(* IEC 61131-3 sources: daoli-st-library/DL_MathData (part 3) *)

(* ---- FC_DL_InterpSegmentWeight.st ---- *)
(*==============================================================================
 * 组件名称 (Component)  : FC_DL_InterpSegmentWeight
 * 所属子库 (Sublibrary) : DL_MathData
 * 当前版本 (Version)    : 1.0.0
 * 兼容性   (Platform)   : CODESYS 3.5+ / TwinCAT 3 / 汇川 InoProShop / 施耐德 Machine Expert
 *                         仅依赖 IEC 61131-3 标准数学（ABS / MIN / MAX），零厂商私有库
 * 功能描述 (Function)   : 段内权重计算：给定升序节点表与查询点，返回相邻两点的
 *                         **加权系数对** (fWLeft, fWRight)，满足 fWLeft + fWRight = 1：
 *                           fWRight = (fXin - afX[i]) / (afX[i+1] - afX[i])
 *                           fWLeft  = 1 - fWRight
 *                         调用方据此自行取 Y（若只有 Y 单表，可算 y = wl*y_i + wr*y_{i+1}），
 *                         也可用于多表共享同一权重（同一 X 上插值多条曲线，
 *                         避免重复定位，性能与一致性双收益）。
 *                         v = wl*v_i + wr*v_{i+1} 与线性插值严格等价（权重和为 1 保证无偏）。
 * 接口     (Interface)  : 输入 afX 升序节点表 [X 单位]、iCount 有效点数 [个]（2..32）、
 *                         fXin 查询点 [X 单位]；
 *                         输出 iSeg 区间左端下标、fWLeft 左节点权重 [0..1]、
 *                         fWRight 右节点权重 [0..1]、bClamped 越界钳位回执、
 *                         eErrCode（E_DL_InterpWgtErr）；
 *                         返回值 = bValid 权重可信标志（TRUE = 两权重可信）。
 * 边界     (Boundary)   : ① 属主边界：只给权重，**不取 Y 值**（取值由调用方组合，
 *                         这是本件与 InterpHoldLast / TwoPointSlope 的本质分工）。
 *                         ② 点数域闸 2..32；越域 → 故障级 eBadCount。
 *                         ③ 非有限双判：查询点 + 全部表元素逐项枚举。
 *                         ④ 段宽近似零 → fWLeft=1.0、fWRight=0.0 并置信息级 eDegenerateSeg
 *                         （权重仍满足和为 1，调用方无需特判；除零被完全规避）。
 *                         ⑤ 越界钳位：fXin 超出 [afX[1], afX[iCount]] → 钳到端段端点，
 *                         权重退化为 (1,0) 或 (0,1)，bClamped=TRUE，不外推。
 *                         ⑥ 权重和复检：|fWLeft + fWRight - 1| < 1E-9，违反 → 故障级 eInternal
 *                         （结构性断言，防未来改动破坏无偏性）。
 *                         ⑦ 零全局耦合（无 GVL / VAR_EXTERNAL / 物理地址）。
 * 分工声明 (Scope)      : 与 `FC_DL_InterpHoldLast` 分工：那件直接给 Y（保持型），
 *                         本件只给权重（多表共享）；与 `FC_DL_TableIndexBinarySearch` 分工：
 *                         大表定位优先用那件，本件为线性扫描 + 权重输出件。
 * 来源标签 (Source Tag) : 原创实现（无外部代码引入）
 * 码表     (Codes)      : 本件不占用全局数字码位；出口为 BOOL + INT + 2×LREAL + BOOL +
 *                         本文件内定义 enum E_DL_InterpWgtErr（全库唯一）。
 * 红线自检 (Redline)    : R1 ✓ 零 GVL/VAR_EXTERNAL ｜ R2 ✓ 零 %I/%Q/%M ｜ R3 ✓ 纯 IEC 61131-3
 *                         R4 ✓ 点数域闸 + 全表非有限双判 + 段宽判零 + 权重和复检 ｜ R5 ✓ 声明逐行同行双语注释
 *                         R6 N/A（纯函数无状态机） ｜ R7 N/A（无实例调用）
 * 修订历史 (Revision)   : 2026-11-23  v1.0.0  R77 首版（批次 B3 · 序号 8）
 * 验收向量 (Acceptance) : ① afX=[0,10,20], iCount=3, fXin=5 → iSeg=1, fWRight=0.5,
 *                         fWLeft=0.5, bClamped=FALSE, eOk, TRUE；
 *                         ② afX 同上, fXin=15 → iSeg=2, fWRight=0.5, fWLeft=0.5；
 *                         ③ afX 同上, fXin=-3 → iSeg=1, fWLeft=1.0, fWRight=0.0, bClamped=TRUE；
 *                         ④ afX 同上, fXin=99 → iSeg=2, fWLeft=0.0, fWRight=1.0, bClamped=TRUE；
 *                         ⑤ afX=[0,0,20], fXin=0 → 退化段：fWLeft=1.0, fWRight=0.0, eDegenerateSeg。
 *==============================================================================*)

(*-----------------------------------------------------------------------------
 * 枚举: E_DL_InterpWgtErr（段内权重错误码，归属 DL_MathData，与本件同文件，全库唯一属主）
 *----------------------------------------------------------------------------*)
TYPE E_DL_InterpWgtErr :
(
    eOk            := 0,   // 信息级：权重计算完成 / Info: weights computed
    eDegenerateSeg := 1,   // 信息级：段宽近似零，权重退化为 1/0 / Info: degenerate segment, weights 1 and 0
    eBadCount      := 2,   // 故障级：点数越域 / Fault: point count out of domain
    eNonFinite     := 3,   // 故障级：查询点或表元素非有限 / Fault: query or table entry non-finite
    eTableNotAsc   := 4,   // 故障级：表不满足升序约定 / Fault: table violates ascending contract
    eInternal      := 9    // 故障级：权重和偏离 1，无偏性被破坏 / Fault: weight sum deviates from one
);
END_TYPE

FUNCTION FC_DL_InterpSegmentWeight : BOOL
VAR_INPUT
    afX    : ARRAY[1..32] OF LREAL;  // 升序节点表 [X 单位] / Ascending node table in X
    iCount : INT;                    // 有效点数（2..32） [个] / Valid point count, 2..32
    fXin   : LREAL;                  // 查询点 [X 单位] / Query value in X
END_VAR
VAR_OUTPUT
    iSeg     : INT;    // 区间左端下标（1..iCount-1） [-] / Segment left index
    fWLeft   : LREAL;  // 左节点权重 [0..1] [-] / Left node weight
    fWRight  : LREAL;  // 右节点权重 [0..1] [-] / Right node weight
    bClamped : BOOL;   // 越界钳位回执 [-] / Out-of-range clamp receipt
    eErrCode : E_DL_InterpWgtErr; // 错误码出口 [-] / Error code outlet
END_VAR
VAR
    _i       : INT;    // 循环下标 [-] / Loop index
    _iSeg    : INT;    // 命中区间下标 [-] / Hit segment index
    _bFound  : BOOL;   // 区间命中标志 [-] / Segment found flag
    _bNonFin : BOOL;   // 非有限标志 [-] / Non-finite flag
    _fDen    : LREAL;  // 段宽（分母） [X 单位] / Segment width denominator
    _fWr     : LREAL;  // 右权重（未钳位） [-] / Raw right weight
    _fSum    : LREAL;  // 权重和（复检用） [-] / Weight sum for recheck
END_VAR
VAR CONSTANT
    DL_IWC_CNT_MIN : INT := 2;        // 点数下限 [个] / Count lower bound
    DL_IWC_CNT_MAX : INT := 32;       // 点数上限（数组容量） [个] / Count upper bound
    DL_IWC_TINY    : LREAL := 1.0E-9; // 段宽近似零阈值 [X 单位] / Degenerate segment threshold
    DL_IWC_ZERO    : LREAL := 0.0;    // 零与权重下限 [-] / Zero and weight lower bound
    DL_IWC_ONE     : LREAL := 1.0;    // 权重上限与无偏基准 [-] / Weight upper bound and unbiasedness base
END_VAR

(* —— 段 0：出口预置安全值（权重预置为「全取左端」，恒满足和为 1） —— *)
FC_DL_InterpSegmentWeight := FALSE;                // 返回值预置无效 / Return preset invalid
iSeg     := 0;                                     // 下标哨兵 / Index sentinel
fWLeft   := DL_IWC_ONE;                            // 左权重哨兵 1（最保守：全取左端） / Left weight sentinel
fWRight  := DL_IWC_ZERO;                           // 右权重哨兵 0 / Right weight sentinel
bClamped := FALSE;                                 // 钳位回执预置否 / Clamp receipt preset false
eErrCode := E_DL_InterpWgtErr.eBadCount;           // 预置最严码 / Preset strictest code

(* —— 段 1：点数域闸 —— *)
IF (iCount < DL_IWC_CNT_MIN) OR (iCount > DL_IWC_CNT_MAX) THEN
    RETURN;
END_IF

(* —— 段 2：非有限域闸（查询点 + 全部表元素逐项枚举） —— *)
_bNonFin := (fXin <> fXin) OR ((fXin - fXin) <> DL_IWC_ZERO);
_i := 1;
WHILE _i <= iCount DO
    IF (afX[_i] <> afX[_i]) OR ((afX[_i] - afX[_i]) <> DL_IWC_ZERO) THEN
        _bNonFin := TRUE;
    END_IF
    _i := _i + 1;
END_WHILE
IF _bNonFin THEN
    eErrCode := E_DL_InterpWgtErr.eNonFinite;
    RETURN;
END_IF

(* —— 段 3：下越界钳位（权重退化 1/0） —— *)
IF fXin <= afX[1] THEN
    iSeg     := 1;
    fWLeft   := DL_IWC_ONE;
    fWRight  := DL_IWC_ZERO;
    bClamped := TRUE;
    eErrCode := E_DL_InterpWgtErr.eOk;
    FC_DL_InterpSegmentWeight := TRUE;
    RETURN;
END_IF

(* —— 段 4：上越界钳位（权重退化 0/1） —— *)
IF fXin >= afX[iCount] THEN
    iSeg     := iCount - 1;
    fWLeft   := DL_IWC_ZERO;
    fWRight  := DL_IWC_ONE;
    bClamped := TRUE;
    eErrCode := E_DL_InterpWgtErr.eOk;
    FC_DL_InterpSegmentWeight := TRUE;
    RETURN;
END_IF

(* —— 段 5：区间定位（升序：afX[i] <= fXin <= afX[i+1]） —— *)
_i      := 1;
_bFound := FALSE;
_iSeg   := 1;
WHILE (_i < iCount) AND (NOT _bFound) DO
    IF (fXin >= afX[_i]) AND (fXin <= afX[_i + 1]) THEN
        _bFound := TRUE;
        _iSeg   := _i;
    ELSE
        _i := _i + 1;
    END_IF
END_WHILE
IF NOT _bFound THEN
    eErrCode := E_DL_InterpWgtErr.eTableNotAsc;    // 未命中：表不升序 / Not found: table not ascending
    RETURN;
END_IF

(* —— 段 6：升序复检 + 段宽判零后计算权重 —— *)
IF afX[_iSeg + 1] < afX[_iSeg] THEN
    eErrCode := E_DL_InterpWgtErr.eTableNotAsc;    // 端点倒序 / Endpoints reversed
    RETURN;
END_IF
_fDen := afX[_iSeg + 1] - afX[_iSeg];              // 段宽 / Segment width
IF ABS(_fDen) < DL_IWC_TINY THEN
    fWLeft   := DL_IWC_ONE;                        // 退化段：全取左端 / Degenerate: all to left
    fWRight  := DL_IWC_ZERO;
    eErrCode := E_DL_InterpWgtErr.eDegenerateSeg;  // 信息级码 / Info code
ELSE
    _fWr     := (fXin - afX[_iSeg]) / _fDen;       // 右权重 / Right weight
    fWRight  := MIN(MAX(_fWr, DL_IWC_ZERO), DL_IWC_ONE);      // 显式约束 0..1 / Constrain 0..1
    fWLeft   := DL_IWC_ONE - fWRight;              // 左权重 = 1 - 右权重（无偏性构造） / Left weight
    eErrCode := E_DL_InterpWgtErr.eOk;             // 信息级成功 / Info success
END_IF
iSeg := _iSeg;

(* —— 段 7：权重和无偏性复检（结构性断言） —— *)
_fSum := fWLeft + fWRight;                         // 权重和 / Weight sum
IF ABS(_fSum - DL_IWC_ONE) > DL_IWC_TINY THEN
    fWLeft   := DL_IWC_ONE;                        // 复检失败：回最保守权重 / Recheck failed: conservative weights
    fWRight  := DL_IWC_ZERO;
    iSeg     := 0;
    eErrCode := E_DL_InterpWgtErr.eInternal;       // 故障级：内部不一致 / Fault: internal inconsistency
    RETURN;
END_IF

FC_DL_InterpSegmentWeight := TRUE;                 // 权重可信 / Weights trustworthy

END_FUNCTION

(* ---- FC_DL_InterpTwoPointSlope.st ---- *)
(*==============================================================================
 * 组件名称 (Component)  : FC_DL_InterpTwoPointSlope
 * 所属子库 (Sublibrary) : DL_MathData
 * 当前版本 (Version)    : 1.0.0
 * 兼容性   (Platform)   : CODESYS 3.5+ / TwinCAT 3 / 汇川 InoProShop / 施耐德 Machine Expert
 *                         仅依赖 IEC 61131-3 标准数学（ABS），零厂商私有库
 * 功能描述 (Function)   : 两点定斜率线性插值 / 受限外推。
 *                           k  = (y2 - y1) / (x2 - x1)                 —— 由两点确定
 *                           y  = y1 + k × (xin - x1)                    —— 通用式（插值外推同一式）
 *                         外推保护：外推距离 = |xin - 近端节点 X|，若超过 fMaxExtrap
 *                         （默认 0.0 = 禁止外推，仅区间内插值），则把 xin 钳到
 *                         「近端节点 ± fMaxExtrap」后再取值，并置 bExtrapolated
 *                         与信息级 eExtrapClamped。**钳位的是 xin 而非 y**，
 *                         这样斜率信息仍可复用（调用方可用 fSlope 自行延续）。
 * 接口     (Interface)  : 输入 fX1/fY1 节点 1、fX2/fY2 节点 2、fXin 查询点、
 *                         fMaxExtrap 允许的最大外推距离 [X 单位，0 = 禁止外推]；
 *                         输出 fYout 结果 [Y 单位]、fSlope 斜率 [Y/X]、
 *                         bExtrapolated 是否发生外推、eErrCode（E_DL_InterpSlopeErr）；
 *                         返回值 = bValid 结果可信标志（TRUE = fYout 可信）。
 * 边界     (Boundary)   : ① 属主边界：只做两点定斜率，不做多点表遍历、不做曲线拟合。
 *                         ② 全浮点入参（7 个）非有限双判，逐一枚举。
 *                         ③ 两点 X 重合（|x2-x1| < 1E-9）→ 故障级 eDegenerateNodes
 *                         （斜率无定义，禁止除零；**先判零后除**）。
 *                         ④ fMaxExtrap < 0 → 故障级 eBadParam（负外推距离无意义）。
 *                         ⑤ fMaxExtrap = 0 表示禁止外推：xin 越界即钳到节点 X，结果 = 端点 Y。
 *                         ⑥ 零全局耦合（无 GVL / VAR_EXTERNAL / 物理地址）。
 * 分工声明 (Scope)      : 与 `FC_DL_InterpLogLinear` 分工：对数域归那件、线性域归本件；
 *                         与 `FC_DL_InterpHoldLast` 分工：保持型（不外推只保持）归那件。
 * 来源标签 (Source Tag) : 原创实现（无外部代码引入）
 * 码表     (Codes)      : 本件不占用全局数字码位；出口为 BOOL + 2×LREAL + BOOL +
 *                         本文件内定义 enum E_DL_InterpSlopeErr（全库唯一）。
 * 红线自检 (Redline)    : R1 ✓ 零 GVL/VAR_EXTERNAL ｜ R2 ✓ 零 %I/%Q/%M ｜ R3 ✓ 纯 IEC 61131-3
 *                         R4 ✓ 全入参非有限双判 + 两点 X 重合判零（除零防护）+ 外推距离上限 ｜ R5 ✓ 声明逐行同行双语注释
 *                         R6 N/A（纯函数无状态机） ｜ R7 N/A（无实例调用）
 * 修订历史 (Revision)   : 2026-11-23  v1.0.0  R77 首版（批次 B3 · 序号 4）
 * 验收向量 (Acceptance) : ① fX1=0, fY1=0, fX2=10, fY2=100, fXin=5, fMaxExtrap=0 → k=10,
 *                         fYout=50.0, bExtrapolated=FALSE, eOk；
 *                         ② 同上, fXin=12, fMaxExtrap=5 → 外推 2 <= 5 → fYout=120.0, eExtrapolated；
 *                         ③ 同上, fXin=20, fMaxExtrap=5 → 钳 xin 到 15 → fYout=150.0, eExtrapClamped；
 *                         ④ fX1=fX2=5 → 返回 FALSE, fYout=0, eDegenerateNodes；
 *                         ⑤ fXin=0, fMaxExtrap=0 → fYout=0.0（左端外推钳到 x1）。
 *==============================================================================*)

(*-----------------------------------------------------------------------------
 * 枚举: E_DL_InterpSlopeErr（两点定斜率插值错误码，归属 DL_MathData，与本件同文件，全库唯一属主）
 *----------------------------------------------------------------------------*)
TYPE E_DL_InterpSlopeErr :
(
    eOk             := 0,   // 信息级：区间内插值 / Info: in-range interpolation
    eExtrapolated   := 1,   // 信息级：受限外推（未超限） / Info: bounded extrapolation within limit
    eExtrapClamped  := 2,   // 信息级：外推超限已钳位 / Info: extrapolation clamped to limit
    eDegenerateNodes:= 3,   // 故障级：两点 X 重合，斜率无定义 / Fault: coincident X, undefined slope
    eBadParam       := 4,   // 故障级：外推距离参数为负 / Fault: negative extrapolation distance
    eNonFinite      := 5    // 故障级：入参非有限 / Fault: non-finite input
);
END_TYPE

FUNCTION FC_DL_InterpTwoPointSlope : BOOL
VAR_INPUT
    fX1        : LREAL;  // 节点 1 的 X [X 单位] / Node one X
    fY1        : LREAL;  // 节点 1 的 Y [Y 单位] / Node one Y
    fX2        : LREAL;  // 节点 2 的 X [X 单位] / Node two X
    fY2        : LREAL;  // 节点 2 的 Y [Y 单位] / Node two Y
    fXin       : LREAL;  // 查询点 X [X 单位] / Query X
    fMaxExtrap : LREAL;  // 允许的最大外推距离（0 = 禁止外推） [X 单位] / Max extrapolation distance, zero forbids
END_VAR
VAR_OUTPUT
    fYout         : LREAL;  // 插值 / 外推结果 [Y 单位] / Interpolated or extrapolated result
    fSlope        : LREAL;  // 两点定出的斜率 [Y/X 单位比] / Slope determined by the two nodes
    bExtrapolated : BOOL;   // 是否发生外推 [-] / Whether extrapolation occurred
    eErrCode      : E_DL_InterpSlopeErr; // 错误码出口 [-] / Error code outlet
END_VAR
VAR
    _bNonFin : BOOL;   // 入参非有限标志 [-] / Non-finite input flag
    _fDx     : LREAL;  // X 方向增量 [X 单位] / X increment
    _fOut    : LREAL;  // 外推距离（带符号） [X 单位] / Signed extrapolation distance
    _fXUse   : LREAL;  // 钳位后实际使用的 X [-] / Actually used X after clamping
    _fLo     : LREAL;  // 允许区间左界 [X 单位] / Allowed lower bound
    _fHi     : LREAL;  // 允许区间右界 [X 单位] / Allowed upper bound
END_VAR
VAR CONSTANT
    DL_ITS_ZERO : LREAL := 0.0;     // 零基准 [-] / Zero base
    DL_ITS_TINY : LREAL := 1.0E-9;  // 两点 X 重合阈值 [X 单位] / Coincident X threshold
END_VAR

(* —— 段 0：出口预置安全值 —— *)
FC_DL_InterpTwoPointSlope := FALSE;                // 返回值预置无效 / Return preset invalid
fYout         := DL_ITS_ZERO;                      // 结果哨兵 0 / Result sentinel
fSlope        := DL_ITS_ZERO;                      // 斜率哨兵 0 / Slope sentinel
bExtrapolated := FALSE;                            // 外推标志预置否 / Extrapolation preset false
eErrCode      := E_DL_InterpSlopeErr.eBadParam;    // 预置最严码 / Preset strictest code

(* —— 段 1：非有限域闸（6 个浮点入参逐一枚举） —— *)
_bNonFin := (fX1 <> fX1) OR ((fX1 - fX1) <> DL_ITS_ZERO);            // X1 非有限 / X1 non-finite
_bNonFin := _bNonFin OR (fY1 <> fY1) OR ((fY1 - fY1) <> DL_ITS_ZERO); // Y1 非有限 / Y1 non-finite
_bNonFin := _bNonFin OR (fX2 <> fX2) OR ((fX2 - fX2) <> DL_ITS_ZERO); // X2 非有限 / X2 non-finite
_bNonFin := _bNonFin OR (fY2 <> fY2) OR ((fY2 - fY2) <> DL_ITS_ZERO); // Y2 非有限 / Y2 non-finite
_bNonFin := _bNonFin OR (fXin <> fXin) OR ((fXin - fXin) <> DL_ITS_ZERO);       // 查询点非有限 / Query non-finite
_bNonFin := _bNonFin OR (fMaxExtrap <> fMaxExtrap) OR ((fMaxExtrap - fMaxExtrap) <> DL_ITS_ZERO); // 外推上限非有限
IF _bNonFin THEN
    eErrCode := E_DL_InterpSlopeErr.eNonFinite;    // 故障级码 / Fault-level code
    RETURN;
END_IF

(* —— 段 2：外推距离参数域闸（不得为负） —— *)
IF fMaxExtrap < DL_ITS_ZERO THEN
    eErrCode := E_DL_InterpSlopeErr.eBadParam;     // 故障级：参数非法 / Fault: illegal parameter
    RETURN;
END_IF

(* —— 段 3：两点 X 重合判零（先判零后做除法，R4 除零防护） —— *)
_fDx := fX2 - fX1;                                 // X 方向增量（分母） / X increment denominator
IF ABS(_fDx) < DL_ITS_TINY THEN
    eErrCode := E_DL_InterpSlopeErr.eDegenerateNodes;  // 故障级：斜率无定义 / Fault: undefined slope
    RETURN;                                        // 早退，杜绝除零 / Early exit, avoids division by zero
END_IF

(* —— 段 4：斜率计算 —— *)
fSlope := (fY2 - fY1) / _fDx;                      // k = dy / dx / Slope

(* —— 段 5：外推距离判定与钳位（钳 xin，不钳 y） —— *)
IF fXin < fX1 THEN
    _fOut := fX1 - fXin;                           // 左向外推距离（正数） / Left extrapolation distance
    IF _fOut > fMaxExtrap THEN
        _fXUse   := fX1 - fMaxExtrap;              // 钳到允许的最远点 / Clamp to farthest allowed point
        eErrCode := E_DL_InterpSlopeErr.eExtrapClamped;   // 信息级：超限钳位 / Info: clamped
    ELSE
        _fXUse   := fXin;                          // 未超限：原值使用 / Within limit: use as-is
        eErrCode := E_DL_InterpSlopeErr.eExtrapolated;    // 信息级：受限外推 / Info: bounded extrapolation
    END_IF
    bExtrapolated := TRUE;                         // 左向外推 / Left extrapolation
ELSIF fXin > fX2 THEN
    _fOut := fXin - fX2;                           // 右向外推距离（正数） / Right extrapolation distance
    IF _fOut > fMaxExtrap THEN
        _fXUse   := fX2 + fMaxExtrap;              // 钳到允许的最远点 / Clamp to farthest allowed point
        eErrCode := E_DL_InterpSlopeErr.eExtrapClamped;   // 信息级：超限钳位 / Info: clamped
    ELSE
        _fXUse   := fXin;                          // 未超限：原值使用 / Within limit: use as-is
        eErrCode := E_DL_InterpSlopeErr.eExtrapolated;    // 信息级：受限外推 / Info: bounded extrapolation
    END_IF
    bExtrapolated := TRUE;                         // 右向外推 / Right extrapolation
ELSE
    _fXUse        := fXin;                         // 区间内插值，无外推 / In-range interpolation
    bExtrapolated := FALSE;
    eErrCode      := E_DL_InterpSlopeErr.eOk;      // 信息级成功 / Info success
END_IF

(* —— 段 6：取值（插值与外推同一式） —— *)
fYout := fY1 + fSlope * (_fXUse - fX1);            // y = y1 + k*(x - x1)

(* —— 段 7：结果非有限复检兜底 —— *)
IF (fYout <> fYout) OR ((fYout - fYout) <> DL_ITS_ZERO) THEN
    fYout         := DL_ITS_ZERO;                  // 复检异常回哨兵 / Recheck failed: sentinel
    fSlope        := DL_ITS_ZERO;
    bExtrapolated := FALSE;
    eErrCode      := E_DL_InterpSlopeErr.eNonFinite;   // 故障级码 / Fault-level code
    RETURN;
END_IF

FC_DL_InterpTwoPointSlope := TRUE;                 // 结果有效 / Result valid

END_FUNCTION

(* ---- FC_DL_IntervalGapCalc.st ---- *)
(*
  ==================================================================
  组件名 Component  : FC_DL_IntervalGapCalc
  分类   Category   : DL_MathData
  前缀   Naming     : FC_DL_ ｜ b/n/u/f/t/e/st 类型前缀制（R265）
  码位   Code ID    : 16#0001_0665（故障级）
  版本   Version    : 1.0.0
  复杂度 Complexity  : 中
  功能   Purpose    : 两区间相离间隙计算：相离返回正间隙宽 [工程单位]，相接 /
                      重叠 / 包含返回 0 并带关系码；供工艺窗对撞分析、换型
                      死区校验、安全包络间距核算等调用方使用。
  开源溯源 Origin    : 西门子 LGF V5.3.0 Comparator 组「区间关系」分类事实
                      借鉴（只借骨不抄肉，与 R11 RangeOverlapCheck 同组既有
                      件互引）；间隙计算 clean-room，零代码复制。
  许可证 License    : MIT
  参考   Reference  : IEC 61131-3:2013 §6.6.1 比较 / MAX 语义
  平台   Platform   : 纯 IEC 61131-3（MAX / ABS / 比较），三平台通用
  依赖   Depends    : 无（零委托、零库件）
  分工声明 Split     : FC_DL_RangeOverlapCheck（五分支关系判定，输出重叠长度）
                      为姊妹件（互引）；本件为「间隙方向」补口：输出相离
                      间隙宽（RangeOverlapCheck 只输出重叠长度，相离时恒 0，
                      间隙量不可观测），两件口径差异显式声明（R216）。
  归属 Ownership     : E_DL_IntervalGap 属主为本文件（全库唯一定义，R264）；
                      引用件只引用不重声明。
  ------------------------------------------------------------------
  边界 Boundary     :
                      一 非有限闸（四个端点 + fEps 逐个点名，R272）：任一
                         非有限 → 故障级 0665 + 返回 eInvalid + fGap = 0 +
                         bValid = FALSE + 早退；
                      二 端点归一：每区间无序端点自动对调，保证下限 ≤ 上限；
                      三 fEps 域闸：负容差非法 → 按默认容差 1.0E-6 接管并
                         并入 0665 处置（与端点非有限出口同形：eInvalid +
                         fGap = 0 + bValid = FALSE，反证句见码表）；
                      四 判定次序写死：相离（正间隙 > fEps）→ 相接（端点
                         重合在容差内）→ 包含 → 部分重叠；相离必须先于
                         相接，相接必须先于重叠（次序不可调换，防多解）；
                      五 完全相等归入 eContained（含端点重合的包含）：相等
                         是包含的退化特例，间隙同为 0，出口无法区分（R90
                         不另立关系码，与 RangeOverlapCheck 的 eEqual 五分
                         支口径差异显式声明）；
                      六 fGap 返回前置非负钳位：舍入产生的微小负值钳到 0；
                      七 纯函数：无记忆量、无定时器、无边沿实例，每调用重算；
                      八 无除法、无循环、无数组访问；无全局、无外部变量、
                         无物理地址。
  错误码 Codes      :
    16#0001_0665【故障级】输入非有限（四端点 / fEps 为 NaN / ±Inf）或 fEps
                         为负（组态非法）
  码位反证 Note     :
    0665 合并「端点 / 容差非有限」与「fEps 为负」的理由：两场景出口组合完全
    相同（eInvalid、fGap = 0、bValid = FALSE、bError = TRUE），三组以内输出
    无法唯一还原该场景，按 R90 不另立码；eInvalid 关系码与 0665 分立：前者
    是返回值语义（关系不可判），后者是诊断码，通道不同不互斥。
  验收 Acceptance   :
    算法已证（脚本）：未跑 ｜ 编译器已证（三平台）：未跑
    V1 相离：A = [0, 10]、B = [20, 30] → eDisjoint、fGap = 10.0
    V2 相接：A = [0, 10]、B = [10, 20] → eTouching、fGap = 0.0
    V3 部分重叠：A = [0, 10]、B = [5, 15] → eOverlap、fGap = 0.0
    V4 包含：A = [0, 10]、B = [2, 8] → eContained、fGap = 0.0
    V5 完全相等：A = B = [0, 10] → eContained（边界五口径）
    V6 无序端点：A = [10, 0] → 归一后同 V1
    V7 端点 NaN → 码 0665 + eInvalid + bValid = FALSE
    V8 fEps = -1.0 → 同码 0665（边界三）
  修订记录 Revision  :
    2026-11-21  v1.0.0  R64 首版（批 1 · 序号 4，LGF Comparator 区间间隙补口）
  ==================================================================
*)
TYPE E_DL_IntervalGap :
(
    eInvalid   := 0,  // 输入非法，关系不可判 / the inputs are illegal, the relation is undecidable
    eDisjoint  := 10, // 完全相离，存在正间隙 / fully disjoint with a positive gap
    eTouching  := 20, // 仅端点相接，间隙为零 / the endpoint touch only with a zero gap
    eOverlap   := 30, // 部分重叠，互不包含 / a partial overlap, neither contains the other
    eContained := 40  // 一方包含另一方（完全相等归入本档）/ one range contains the other, an equality is folded here
);
END_TYPE

FUNCTION FC_DL_IntervalGapCalc : E_DL_IntervalGap
VAR_INPUT
    fA1  : LREAL := 0.0;    // 区间 A 端点 1 [工程单位]，无序自动对调 / the range A endpoint one, auto swapped
    fA2  : LREAL := 10.0;   // 区间 A 端点 2 [工程单位] / the range A endpoint two
    fB1  : LREAL := 0.0;    // 区间 B 端点 1 [工程单位]，无序自动对调 / the range B endpoint one, auto swapped
    fB2  : LREAL := 10.0;   // 区间 B 端点 2 [工程单位] / the range B endpoint two
    fEps : LREAL := 1.0E-6; // 容差 [工程单位]，≥ 0 / the tolerance, non negative
END_VAR
VAR_OUTPUT
    fGap   : LREAL; // 相离间隙宽 [工程单位]，恒非负，非相离 = 0.0 / the gap width, never negative, zero unless disjoint
    bValid : BOOL;  // 结果可用 [-] / the result usable flag
    eErr   : UDINT; // 错误码，0 = 正常 / the error code, zero is ok
    bError : BOOL;  // 故障标志（故障级码同拍置位，R45 配对）/ the fault flag raised with a fault level code
END_VAR
VAR
    _fLoA   : LREAL := 0.0; // 区间 A 归一下限 [工程单位] / the normalised lower bound of the range A
    _fHiA   : LREAL := 0.0; // 区间 A 归一上限 [工程单位] / the normalised upper bound of the range A
    _fLoB   : LREAL := 0.0; // 区间 B 归一下限 [工程单位] / the normalised lower bound of the range B
    _fHiB   : LREAL := 0.0; // 区间 B 归一上限 [工程单位] / the normalised upper bound of the range B
    _fTmp   : LREAL := 0.0; // 对调临时量 [工程单位] / the swap temporary
    _fGapUse: LREAL := 0.0; // 间隙工作副本 [工程单位] / the gap working copy
    _fEpsUse: LREAL := 0.0; // 容差工作副本 [工程单位] / the tolerance working copy
END_VAR  // R64 结构补齐：VAR 段缺失的 END_VAR（门禁机械修复）
VAR CONSTANT
    DL_IGP_ZERO : LREAL := 0.0;    // 实数零常量 [工程单位] / the real zero constant
    DL_IGP_EPSDF: LREAL := 1.0E-6; // 默认容差常量 [工程单位]（fEps 非法时接管）/ the default tolerance taken over when the input is illegal
END_VAR

// 段 1｜返回值与全部出口预置安全值（R45 四段式第一段）/ segment 1, the preset of the return and all outlets
FC_DL_IntervalGapCalc := E_DL_IntervalGap.eInvalid; // 返回值预置不可判（任何早退天然带不可判语义）/ preset the return to undecidable
fGap := DL_IGP_ZERO; // 间隙预置零 [工程单位] / preset the gap zero
bValid := FALSE; // 可用标志预置假 / preset the validity false
eErr := 16#0000_0000; // 错误码预置正常 / preset the code to ok
bError := FALSE; // 故障标志预置假 / preset the fault flag false
_fLoA := DL_IGP_ZERO; // 归一下限 A 预置零 / preset the lower bound A zero
_fHiA := DL_IGP_ZERO; // 归一上限 A 预置零 / preset the upper bound A zero
_fLoB := DL_IGP_ZERO; // 归一下限 B 预置零 / preset the lower bound B zero
_fHiB := DL_IGP_ZERO; // 归一上限 B 预置零 / preset the upper bound B zero
_fTmp := DL_IGP_ZERO; // 对调临时量预置零 / preset the swap temporary zero
_fGapUse := DL_IGP_ZERO; // 间隙工作副本预置零 / preset the gap copy zero
_fEpsUse := DL_IGP_EPSDF; // 容差工作副本预置默认容差 / preset the tolerance copy to the default

// 段 2｜非有限闸与容差域闸（边界一 / 边界三，逐个点名，R272）/ segment 2, the finiteness gate and the tolerance gate
IF (fA1 <> fA1) OR ((fA1 - fA1) <> (fA1 - fA1))
OR (fA2 <> fA2) OR ((fA2 - fA2) <> (fA2 - fA2))
OR (fB1 <> fB1) OR ((fB1 - fB1) <> (fB1 - fB1))
OR (fB2 <> fB2) OR ((fB2 - fB2) <> (fB2 - fB2))
OR (fEps <> fEps) OR ((fEps - fEps) <> (fEps - fEps))
OR (fEps < DL_IGP_ZERO) THEN // 任一端点 / 容差非有限或容差为负 / any endpoint or the tolerance is not finite or negative
    eErr := 16#0001_0665; // 故障级：输入非有限或容差非法（出口同形合并一码，R90）/ fault grade under the merged code
    bError := TRUE; // 同拍置故障标志（R45 配对）/ raise the fault flag on the same scan
    bValid := FALSE; // 结果不可用 / the result is not usable
    RETURN; // 早退，返回 eInvalid / early return with undecidable
END_IF
_fEpsUse := fEps; // 容差接管（已证非负有限）[工程单位] / take the tolerance proven nonnegative and finite

// 段 3｜端点归一（边界二：无序端点自动对调）/ segment 3, the endpoint normalisation with the auto swap
_fLoA := fA1; // A 下限暂存端点 1 / the A lower takes the endpoint one
_fHiA := fA2; // A 上限暂存端点 2 / the A upper takes the endpoint two
IF _fLoA > _fHiA THEN // A 端点逆序 / the A endpoints in reverse order
    _fTmp := _fLoA; // 暂存下限 / save the lower
    _fLoA := _fHiA; // 下限取原上限 / the lower takes the former upper
    _fHiA := _fTmp; // 上限取原下限 / the upper takes the former lower
END_IF
_fLoB := fB1; // B 下限暂存端点 1 / the B lower takes the endpoint one
_fHiB := fB2; // B 上限暂存端点 2 / the B upper takes the endpoint two
IF _fLoB > _fHiB THEN // B 端点逆序 / the B endpoints in reverse order
    _fTmp := _fLoB; // 暂存下限 / save the lower
    _fLoB := _fHiB; // 下限取原上限 / the lower takes the former upper
    _fHiB := _fTmp; // 上限取原下限 / the upper takes the former lower
END_IF

// 段 4｜关系与间隙判定（边界四：次序写死，相离 → 相接 → 包含 → 重叠）/ segment 4, the relation and gap in the frozen order
IF (_fLoB - _fHiA) > _fEpsUse THEN // B 整体在 A 右侧且存在正间隙 / the B sits right with a positive gap
    _fGapUse := _fLoB - _fHiA; // 间隙 = B 下限 − A 上限 [工程单位] / the gap of the B lower minus the A upper
    FC_DL_IntervalGapCalc := E_DL_IntervalGap.eDisjoint; // 相离关系 / the disjoint relation
ELSIF (_fLoA - _fHiB) > _fEpsUse THEN // A 整体在 B 右侧且存在正间隙 / the A sits right with a positive gap
    _fGapUse := _fLoA - _fHiB; // 间隙 = A 下限 − B 上限 [工程单位] / the gap of the A lower minus the B upper
    FC_DL_IntervalGapCalc := E_DL_IntervalGap.eDisjoint; // 相离关系 / the disjoint relation
ELSIF (ABS(_fHiA - _fLoB) < _fEpsUse) OR (ABS(_fHiB - _fLoA) < _fEpsUse) THEN // 端点几何重合（容差内）/ the endpoints coincide inside the tolerance
    _fGapUse := DL_IGP_ZERO; // 相接间隙为零 [工程单位] / the touching gap zero
    FC_DL_IntervalGapCalc := E_DL_IntervalGap.eTouching; // 相接关系 / the touching relation
ELSIF ((_fLoA <= _fLoB + _fEpsUse) AND (_fHiA >= _fHiB - _fEpsUse))
OR ((_fLoB <= _fLoA + _fEpsUse) AND (_fHiB >= _fHiA - _fEpsUse)) THEN // 一方包含另一方（含完全相等退化特例，边界五）/ one contains the other, an equality folded in
    _fGapUse := DL_IGP_ZERO; // 包含间隙为零 [工程单位] / the contained gap zero
    FC_DL_IntervalGapCalc := E_DL_IntervalGap.eContained; // 包含关系 / the contained relation
ELSE // 部分重叠（互不包含，间隙恒 0）/ a partial overlap with a zero gap
    _fGapUse := DL_IGP_ZERO; // 重叠间隙为零 [工程单位] / the overlap gap zero
    FC_DL_IntervalGapCalc := E_DL_IntervalGap.eOverlap; // 部分重叠关系 / the partial overlap relation
END_IF

// 段 5｜间隙非负钳位与统一出口（边界六）/ segment 5, the nonnegative clamp and the unified outlet
IF _fGapUse < DL_IGP_ZERO THEN // 舍入产生微小负值 / a tiny negative from the rounding
    _fGapUse := DL_IGP_ZERO; // 钳到 0，维持非负承诺 / clamp to zero, keep the promise
END_IF
fGap := _fGapUse; // 间隙出口 [工程单位] / the gap outlet
bValid := TRUE; // 结果可用 / the result is usable
END_FUNCTION

(* ---- FC_DL_LengthUnitConvert.st ---- *)
(*==============================================================================
 * 组件名称 (Component)  : FC_DL_LengthUnitConvert
 * 所属子库 (Sublibrary) : DL_MathData
 * 当前版本 (Version)    : 1.0.0
 * 兼容性   (Platform)   : CODESYS 3.5+ / TwinCAT 3 / 汇川 InoProShop / 施耐德 Machine Expert
 *                         仅依赖 IEC 61131-3 算术运算符，零厂商私有库
 * 功能描述 (Function)   : 长度工程量单位换算（系数表驱动）：以米（m）为中介单位，
 *                         fHub = fValue × kSrc，fResult = fHub ÷ kDst；
 *                         kSrc / kDst 为编译期非零常量，纯常量除法，结构性无除零。
 *                         长度物理量非负：负值判故障级 eNegativeValue 并回哨兵 0；
 *                         零值合法（0 mm = 0 m，info 级 eZeroValue）。
 * 接口     (Interface)  : 输入 fValue 被换算长度 [源单位]、eSrc 源单位、eDst 目标单位；
 *                         输出 fConverted 换算结果 [目标单位]、eErrCode 错误码（E_DL_LenConvErr）；
 *                         返回值 = bValid 数值可信标志（TRUE = fConverted 可信）。
 * 边界     (Boundary)   : ① 属主边界：只做单位换算，不做量程标定、不做累计行程管理。
 *                         ② 单位枚举越域（非四成员之一）→ 故障级 eInvalidUnit，结果哨兵 0。
 *                         ③ 全浮点入参做非有限双判（NaN 自反 / Inf 差自减），任一非有限 →
 *                         故障级 eNonFinite。中介值与结果各复检一次（四段式第四段）。
 *                         ④ 负长度 → 故障级 eNegativeValue（物理量不可为负，拒绝换算而非钳位，
 *                         避免掩盖上游符号错误）。钳位会静默改值，故不采用。
 *                         ⑤ 零全局耦合（无 GVL / VAR_EXTERNAL / 物理地址）。
 * 分工声明 (Scope)      : 与 `FC_DL_PressUnitConvert` 同族不同量（压力含负压域、长度不含）；
 *                         与 `FC_DL_AreaUnitConvert` 分工：长度 ↔ 面积不做隐式平方推导。
 * 来源标签 (Source Tag) : 开源溯源：lgf-math 换算系数（公开物理常数，clean-room 重写）；许可证 MIT（仅参考语义，代码原创）
 * 码表     (Codes)      : 本件不占用全局数字码位；出口为 BOOL + LREAL + 本文件内定义
 *                         enum E_DL_LenConvErr（全库唯一）。
 * 红线自检 (Redline)    : R1 ✓ 零 GVL/VAR_EXTERNAL ｜ R2 ✓ 零 %I/%Q/%M ｜ R3 ✓ 纯 IEC 61131-3
 *                         R4 ✓ 非有限双判 + 枚举域闸 + 常量除法无除零 + 负值拒绝 ｜ R5 ✓ 声明逐行同行双语注释
 *                         R6 N/A（纯函数无状态机） ｜ R7 N/A（无实例调用）
 * 修订历史 (Revision)   : 2026-11-23  v1.0.0  R77 首版（批次 B2 · 序号 11）
 * 验收向量 (Acceptance) : ① fValue=1000, eSrc=eMm, eDst=eM → 1000×0.001 = 1.0 m, eOk, TRUE；
 *                         ② fValue=1.0, eSrc=eInch, eDst=eMm → 1×0.0254 = 0.0254 m,
 *                         ÷0.001 = 25.4 mm（容差 1E-9）；
 *                         ③ fValue=1.0, eSrc=eFt, eDst=eM → 0.3048 m, eOk；
 *                         ④ fValue=-5.0, eSrc=eMm, eDst=eM → 返回 FALSE, fConverted=0, eNegativeValue；
 *                         ⑤ fValue=0.0, eSrc=eMm, eDst=eFt → 0.0, 返回 TRUE, eZeroValue。
 *==============================================================================*)

(*-----------------------------------------------------------------------------
 * 枚举: E_DL_LengthUnit（长度单位表，归属 DL_MathData，与本件同文件，全库唯一属主）
 *----------------------------------------------------------------------------*)
TYPE E_DL_LengthUnit :
(
    eMm   := 0,   // 毫米（中介单位 m 的千分之一） / Millimetre, one thousandth of hub metre
    eM    := 1,   // 米（中介单位） / Metre, hub unit
    eInch := 2,   // 英寸（25.4 mm） / Inch, exactly 25.4 mm
    eFt   := 3    // 英尺（12 英寸） / Foot, twelve inches
);
END_TYPE

(*-----------------------------------------------------------------------------
 * 枚举: E_DL_LenConvErr（长度换算错误码）
 * 分级: eNegativeValue / eInvalidUnit / eNonFinite 为故障级（返回 FALSE）；
 *       eOk / eZeroValue 为信息级（返回 TRUE）。
 *----------------------------------------------------------------------------*)
TYPE E_DL_LenConvErr :
(
    eOk            := 0,   // 信息级：换算完成 / Info: conversion completed
    eZeroValue     := 1,   // 信息级：输入为零（合法） / Info: zero input, legal
    eInvalidUnit   := 2,   // 故障级：单位枚举越域 / Fault: unit enum out of domain
    eNonFinite     := 3,   // 故障级：输入非有限 / Fault: non-finite input
    eNegativeValue := 4    // 故障级：负长度 / Fault: negative length
);
END_TYPE

FUNCTION FC_DL_LengthUnitConvert : BOOL
VAR_INPUT
    fValue : LREAL;            // 被换算长度值 [源单位] / Length value in source unit
    eSrc   : E_DL_LengthUnit;  // 源单位枚举 [-] / Source unit enum
    eDst   : E_DL_LengthUnit;  // 目标单位枚举 [-] / Destination unit enum
END_VAR
VAR_OUTPUT
    fConverted : LREAL;            // 换算结果 [目标单位] / Converted result in destination unit
    eErrCode   : E_DL_LenConvErr;  // 错误码出口 [-] / Error code outlet
END_VAR
VAR
    _bNonFin : BOOL;   // 输入非有限当拍标志 [-] / Non-finite input flag
    _fHub    : LREAL;  // 中介长度值 [m] / Hub length value in metres
END_VAR
VAR CONSTANT
    DL_LUC_MM   : LREAL := 0.001;    // mm → m 换算系数 [m/mm] / mm to m factor
    DL_LUC_M    : LREAL := 1.0;      // m → m 恒等系数 [m/m] / m identity factor
    DL_LUC_INCH : LREAL := 0.0254;   // inch → m 换算系数 [m/inch] / inch to m factor
    DL_LUC_FT   : LREAL := 0.3048;   // ft → m 换算系数 [m/ft] / foot to m factor
    DL_LUC_ZERO : LREAL := 0.0;      // 零值与非有限判零基准 [-] / Zero and non-finite base
END_VAR

(* —— 段 0：出口预置安全值 —— *)
FC_DL_LengthUnitConvert := FALSE;                  // 返回值预置无效 / Return preset invalid
fConverted := DL_LUC_ZERO;                         // 结果哨兵 0 / Result sentinel zero
eErrCode   := E_DL_LenConvErr.eInvalidUnit;        // 预置最严码 / Preset strictest code

(* —— 段 1：非有限域闸（R79 双判：NaN 自反 + Inf 差自减） —— *)
_bNonFin := (fValue <> fValue) OR ((fValue - fValue) <> DL_LUC_ZERO);   // 非有限判定 / Non-finite test
IF _bNonFin THEN
    eErrCode := E_DL_LenConvErr.eNonFinite;        // 故障级码 / Fault-level code
    RETURN;                                        // 早退保持哨兵 / Early exit with sentinel
END_IF

(* —— 段 2：负长度域闸（物理量不可为负，拒绝而非钳位） —— *)
IF fValue < DL_LUC_ZERO THEN
    eErrCode := E_DL_LenConvErr.eNegativeValue;    // 故障级码 / Fault-level code
    RETURN;                                        // 早退保持哨兵 / Early exit with sentinel
END_IF

(* —— 段 3：源单位 → 中介米（按枚举成员逐值比较，不依赖 ENUM→INT 强转方言） —— *)
IF eSrc = E_DL_LengthUnit.eMm THEN
    _fHub := fValue * DL_LUC_MM;                   // mm × 0.001 / mm scaled
ELSIF eSrc = E_DL_LengthUnit.eM THEN
    _fHub := fValue * DL_LUC_M;                    // m 直通 / metre pass-through
ELSIF eSrc = E_DL_LengthUnit.eInch THEN
    _fHub := fValue * DL_LUC_INCH;                 // inch × 0.0254 / inch scaled
ELSIF eSrc = E_DL_LengthUnit.eFt THEN
    _fHub := fValue * DL_LUC_FT;                   // ft × 0.3048 / foot scaled
ELSE
    RETURN;                                        // 源单位越域：保持预置故障码 / Source unit out of domain
END_IF

(* —— 段 4：中介米 → 目标单位（常量除法，分母非零结构性无除零） —— *)
IF eDst = E_DL_LengthUnit.eMm THEN
    fConverted := _fHub / DL_LUC_MM;               // ÷0.001 / Divide by mm factor
ELSIF eDst = E_DL_LengthUnit.eM THEN
    fConverted := _fHub / DL_LUC_M;                // ÷1 / Divide by identity
ELSIF eDst = E_DL_LengthUnit.eInch THEN
    fConverted := _fHub / DL_LUC_INCH;             // ÷0.0254 / Divide by inch factor
ELSIF eDst = E_DL_LengthUnit.eFt THEN
    fConverted := _fHub / DL_LUC_FT;               // ÷0.3048 / Divide by foot factor
ELSE
    eErrCode   := E_DL_LenConvErr.eInvalidUnit;    // 目标单位越域 / Destination unit out of domain
    fConverted := DL_LUC_ZERO;                     // 结果回哨兵 / Result back to sentinel
    RETURN;                                        // 早退 / Early exit
END_IF

(* —— 段 5：结果非有限复检兜底（四段式第四段） —— *)
IF (fConverted <> fConverted) OR ((fConverted - fConverted) <> DL_LUC_ZERO) THEN
    fConverted := DL_LUC_ZERO;                     // 复检异常回哨兵 / Recheck failed: sentinel
    eErrCode   := E_DL_LenConvErr.eNonFinite;      // 故障级码 / Fault-level code
    RETURN;                                        // 早退 / Early exit
END_IF

(* —— 段 6：成功出口（零值单独置信息码，仍算有效换算） —— *)
IF fValue = DL_LUC_ZERO THEN
    eErrCode := E_DL_LenConvErr.eZeroValue;        // 信息级：零值 / Info: zero value
ELSE
    eErrCode := E_DL_LenConvErr.eOk;               // 信息级成功 / Info success
END_IF
FC_DL_LengthUnitConvert := TRUE;                   // 换算有效 / Conversion valid

END_FUNCTION

(* ---- FC_DL_MassUnitConvert.st ---- *)
(*==============================================================================
 * 组件名称 (Component)  : FC_DL_MassUnitConvert
 * 所属子库 (Sublibrary) : DL_MathData
 * 当前版本 (Version)    : 1.0.0
 * 兼容性   (Platform)   : CODESYS 3.5+ / TwinCAT 3 / 汇川 InoProShop / 施耐德 Machine Expert
 *                         仅依赖 IEC 61131-3 算术运算符，零厂商私有库
 * 功能描述 (Function)   : 质量工程量单位换算（系数表驱动）：以千克（kg）为中介单位，
 *                         fHub = fValue × kSrc，fResult = fHub ÷ kDst；系数为编译期
 *                         非零常量，纯常量除法，结构性无除零。
 *                         质量非负：负值判故障级 eNegativeValue 并回哨兵 0（称重去皮负数
 *                         属上游补偿问题，必须显式拒绝，禁止在此静默取绝对值）。
 * 接口     (Interface)  : 输入 fValue 被换算质量 [源单位]、eSrc 源单位、eDst 目标单位；
 *                         输出 fConverted 换算结果 [目标单位]、eErrCode（E_DL_MassConvErr）；
 *                         返回值 = bValid 数值可信标志（TRUE = fConverted 可信）。
 * 边界     (Boundary)   : ① 属主边界：只做单位换算，不做去皮 / 标定 / 累计称重。
 *                         ② 单位枚举越域 → 故障级 eInvalidUnit，结果哨兵 0。
 *                         ③ 非有限双判（NaN 自反 / Inf 差自减），命中即故障级 eNonFinite。
 *                         ④ 负质量 → 故障级 eNegativeValue（拒绝换算，不钳位）。
 *                         ⑤ 零值合法（info 级 eZeroValue）。结果与中介值各复检一次。
 *                         ⑥ 零全局耦合（无 GVL / VAR_EXTERNAL / 物理地址）。
 * 分工声明 (Scope)      : 与 `FC_DL_LengthUnitConvert` 同族不同量；与称重 FB 分工：
 *                         重量采集与稳定判据归称重 FB，本件只做单位间换算。
 * 来源标签 (Source Tag) : 开源溯源：lgf-math 换算系数（公开物理常数，clean-room 重写）；许可证 MIT（仅参考语义，代码原创）
 * 码表     (Codes)      : 本件不占用全局数字码位；出口为 BOOL + LREAL +
 *                         本文件内定义 enum E_DL_MassConvErr（全库唯一）。
 * 红线自检 (Redline)    : R1 ✓ 零 GVL/VAR_EXTERNAL ｜ R2 ✓ 零 %I/%Q/%M ｜ R3 ✓ 纯 IEC 61131-3
 *                         R4 ✓ 非有限双判 + 枚举域闸 + 常量除法无除零 + 负值拒绝 ｜ R5 ✓ 声明逐行同行双语注释
 *                         R6 N/A（纯函数无状态机） ｜ R7 N/A（无实例调用）
 * 修订历史 (Revision)   : 2026-11-23  v1.0.0  R77 首版（批次 B2 · 序号 12）
 * 验收向量 (Acceptance) : ① fValue=1000, eSrc=eG, eDst=eKg → 1000×0.001 = 1.0 kg, eOk, TRUE；
 *                         ② fValue=1.0, eSrc=eLb, eDst=eG → 1×0.45359237 = 0.45359237 kg,
 *                         ÷0.001 = 453.59237 g（容差 1E-9）；
 *                         ③ fValue=16.0, eSrc=eOz, eDst=eLb → 16×0.028349523125 =
 *                         0.45359237 kg, ÷0.45359237 = 1.0 lb（容差 1E-9）；
 *                         ④ fValue=-1.0, eSrc=eKg, eDst=eG → 返回 FALSE, 0, eNegativeValue。
 *==============================================================================*)

(*-----------------------------------------------------------------------------
 * 枚举: E_DL_MassUnit（质量单位表，归属 DL_MathData，与本件同文件，全库唯一属主）
 *----------------------------------------------------------------------------*)
TYPE E_DL_MassUnit :
(
    eG  := 0,   // 克（中介单位 kg 的千分之一） / Gram, one thousandth of hub kilogram
    eKg := 1,   // 千克（中介单位） / Kilogram, hub unit
    eLb := 2,   // 磅（常衡，0.45359237 kg） / Pound avoirdupois
    eOz := 3    // 盎司（常衡，1/16 磅） / Ounce avoirdupois, one sixteenth of pound
);
END_TYPE

(*-----------------------------------------------------------------------------
 * 枚举: E_DL_MassConvErr（质量换算错误码）
 *----------------------------------------------------------------------------*)
TYPE E_DL_MassConvErr :
(
    eOk            := 0,   // 信息级：换算完成 / Info: conversion completed
    eZeroValue     := 1,   // 信息级：输入为零（合法） / Info: zero input, legal
    eInvalidUnit   := 2,   // 故障级：单位枚举越域 / Fault: unit enum out of domain
    eNonFinite     := 3,   // 故障级：输入非有限 / Fault: non-finite input
    eNegativeValue := 4    // 故障级：负质量 / Fault: negative mass
);
END_TYPE

FUNCTION FC_DL_MassUnitConvert : BOOL
VAR_INPUT
    fValue : LREAL;          // 被换算质量值 [源单位] / Mass value in source unit
    eSrc   : E_DL_MassUnit;  // 源单位枚举 [-] / Source unit enum
    eDst   : E_DL_MassUnit;  // 目标单位枚举 [-] / Destination unit enum
END_VAR
VAR_OUTPUT
    fConverted : LREAL;            // 换算结果 [目标单位] / Converted result
    eErrCode   : E_DL_MassConvErr; // 错误码出口 [-] / Error code outlet
END_VAR
VAR
    _bNonFin : BOOL;   // 输入非有限当拍标志 [-] / Non-finite input flag
    _fHub    : LREAL;  // 中介质量值 [kg] / Hub mass value in kilograms
END_VAR
VAR CONSTANT
    DL_MUC_G    : LREAL := 0.001;           // g → kg 换算系数 [kg/g] / gram to kilogram factor
    DL_MUC_KG   : LREAL := 1.0;             // kg → kg 恒等系数 [kg/kg] / kilogram identity factor
    DL_MUC_LB   : LREAL := 0.45359237;      // lb → kg 换算系数（常衡精确定义） [kg/lb] / pound to kilogram factor
    DL_MUC_OZ   : LREAL := 0.028349523125;  // oz → kg 换算系数（lb/16） [kg/oz] / ounce to kilogram factor
    DL_MUC_ZERO : LREAL := 0.0;             // 零值与非有限判零基准 [-] / Zero and non-finite base
END_VAR

(* —— 段 0：出口预置安全值 —— *)
FC_DL_MassUnitConvert := FALSE;                    // 返回值预置无效 / Return preset invalid
fConverted := DL_MUC_ZERO;                         // 结果哨兵 0 / Result sentinel
eErrCode   := E_DL_MassConvErr.eInvalidUnit;       // 预置最严码 / Preset strictest code

(* —— 段 1：非有限域闸（R79 双判） —— *)
_bNonFin := (fValue <> fValue) OR ((fValue - fValue) <> DL_MUC_ZERO);   // 非有限判定 / Non-finite test
IF _bNonFin THEN
    eErrCode := E_DL_MassConvErr.eNonFinite;       // 故障级码 / Fault-level code
    RETURN;
END_IF

(* —— 段 2：负质量域闸（拒绝换算，不静默取绝对值） —— *)
IF fValue < DL_MUC_ZERO THEN
    eErrCode := E_DL_MassConvErr.eNegativeValue;   // 故障级码 / Fault-level code
    RETURN;
END_IF

(* —— 段 3：源单位 → 中介千克 —— *)
IF eSrc = E_DL_MassUnit.eG THEN
    _fHub := fValue * DL_MUC_G;                    // g × 0.001 / gram scaled
ELSIF eSrc = E_DL_MassUnit.eKg THEN
    _fHub := fValue * DL_MUC_KG;                   // kg 直通 / kilogram pass-through
ELSIF eSrc = E_DL_MassUnit.eLb THEN
    _fHub := fValue * DL_MUC_LB;                   // lb × 0.45359237 / pound scaled
ELSIF eSrc = E_DL_MassUnit.eOz THEN
    _fHub := fValue * DL_MUC_OZ;                   // oz × 0.028349523125 / ounce scaled
ELSE
    RETURN;                                        // 源单位越域 / Source unit out of domain
END_IF

(* —— 段 4：中介千克 → 目标单位（常量除法，分母非零） —— *)
IF eDst = E_DL_MassUnit.eG THEN
    fConverted := _fHub / DL_MUC_G;                // ÷0.001 / Divide by gram factor
ELSIF eDst = E_DL_MassUnit.eKg THEN
    fConverted := _fHub / DL_MUC_KG;               // ÷1 / Divide by identity
ELSIF eDst = E_DL_MassUnit.eLb THEN
    fConverted := _fHub / DL_MUC_LB;               // ÷0.45359237 / Divide by pound factor
ELSIF eDst = E_DL_MassUnit.eOz THEN
    fConverted := _fHub / DL_MUC_OZ;               // ÷0.028349523125 / Divide by ounce factor
ELSE
    eErrCode   := E_DL_MassConvErr.eInvalidUnit;   // 目标单位越域 / Destination out of domain
    fConverted := DL_MUC_ZERO;
    RETURN;
END_IF

(* —— 段 5：结果非有限复检兜底 —— *)
IF (fConverted <> fConverted) OR ((fConverted - fConverted) <> DL_MUC_ZERO) THEN
    fConverted := DL_MUC_ZERO;                     // 复检异常回哨兵 / Recheck failed: sentinel
    eErrCode   := E_DL_MassConvErr.eNonFinite;     // 故障级码 / Fault-level code
    RETURN;
END_IF

(* —— 段 6：成功出口 —— *)
IF fValue = DL_MUC_ZERO THEN
    eErrCode := E_DL_MassConvErr.eZeroValue;       // 信息级：零值 / Info: zero value
ELSE
    eErrCode := E_DL_MassConvErr.eOk;              // 信息级成功 / Info success
END_IF
FC_DL_MassUnitConvert := TRUE;                     // 换算有效 / Conversion valid

END_FUNCTION

(* ---- FC_DL_ModbusExceptionParse.st ---- *)
(*==============================================================================
 * 组件名称 (Component)  : FC_DL_ModbusExceptionParse
 * 所属子库 (Sublibrary) : DL_MathData
 * 归属目录 (Directory)  : C:\Library\DL_MathData
 * 当前版本 (Version)    : 1.0.0
 * 组件分类 (Category)   : 函数（FUNCTION）· 纯函数 · 协议诊断帧解析
 * 兼容性   (Platform)   : CODESYS 3.5 / TwinCAT 3 / 汇川 InoProShop / 施耐德
 *                         Machine Expert；仅用标准位运算与枚举，无实例依赖
 * 功能一句话 (Summary)  : 解析从站异常响应帧（功能码最高位置位加异常码），输出原始
 *                         功能码、异常码中文名、严重度分级与可重试标志。
 * 功能描述 (Function)   : 从站回非法数据地址与回从站设备忙，在通讯层都只表现为
 *                         「事务失败」；前者是组态错必须改程序，后者重试即可。
 *                         现场一律当「通讯不稳」处理，反复重启总线。本件把两者
 *                         分开定性，让上层重试策略按严重度分级动作。
 * 与既有件边界 (Boundary): FB_DL_ModbusPollMaster 负责组帧、发送、超时与重试编排；
 *                         本件只解析不决策，是否重试、重试几次由调用方的重试上限
 *                         决定。二者是「判读」与「执行」的分工，本件不持有任何状态。
 * 设计要点 (Key notes)  : ① 功能码先去最高位得原始码，原始码为零视为帧不可解释；
 *                         ② 非异常帧也走完整出口，返回「正常响应」文字与信息码，
 *                           便于 HMI 用同一字段显示两种帧；
 *                         ③ 未定义异常码不算解析成功：文字照给，但有效性置假，
 *                           让上层既能显示又能区分「看不懂」与「看懂且是故障」；
 *                         ④ 严重度分级是本件的核心输出，重试判据与分级绑定，
 *                           避免上层拿「故障」去无脑重试；
 *                         ⑤ 纯函数：无算术、无除法、无循环、无内部状态。
 * 开源溯源 (Origin)     : 来源标签 oscat-network。OSCAT 为公开发布的第三方函数库，
 *                         本件仅借鉴其把「协议帧解析 / 校验 / 诊断」分成独立函数族
 *                         的分类方式，以及「功能码 + 异常码」两入参的参数域；许可证
 *                         按其发布方条款仅作分类参考，本件零代码行、零注释引用。
 *                         异常码语义取自 Modbus 应用协议规范的公开定义（该规范为公开
 *                         技术文档），中文名、分级与可重试判据为本库自有设计，
 *                         整体属 clean-room 独立实现。
 * 码位说明 (Codes)      : 本件独占信息级码段 16#0001_0138 到 16#0001_0139，纯函数
 *                         无锁存面故不占故障级码；与同族 0134 到 013C 各件相邻不重叠。
 *                         0138 功能码非法或异常码未定义 ｜ 0139 本帧非异常帧。
 * 依赖说明 (Depends)    : 无 DL_ 内部依赖；仅 Standard.library 的位运算与
 *                         USINT_TO_INT 显式转换。
 * 红线自检 (Redline)    : 零全局变量表依赖 ｜ 零外部变量声明 ｜ 零物理地址
 *                         纯 IEC 61131-3 ｜ 无算术无除法 ｜ 分支带兜底
 *                         全变量双语同行注释 ｜ 无定时器实例
 * 修订历史 (Revision)   : 2026-11-15  v1.0.0  首版入库（Round 12 · 协议诊断族）
 *============================================================================*)

(*-----------------------------------------------------------------------------
 * 枚举: E_DL_ModbusExcSeverity（归属 DL_MathData，与本件同文件）
 * 含义: 异常码的处置严重度。编号 0 起跳、段间隔 10。
 *----------------------------------------------------------------------------*)
TYPE E_DL_ModbusExcSeverity :
(
    eInfo  := 0,     // 提示级：可忽略，不改变重试策略 / Informational, no retry impact
    eWarn  := 10,    // 告警级：可原样重试，短退避后再发 / Warning, safe to retry after a short back off
    eFault := 20     // 故障级：须人工介入，重试无意义或有害 / Fault, manual intervention required
);
END_TYPE

(*==============================================================================
 * 判读示意 (Interpretation picture)：
 *   功能码 16#83 表示读保持寄存器出错，去掉最高位得原始码 3
 *   异常码 16#02 语义为非法数据地址，属组态错，故障级，不可重试
 *   功能码 16#86 表示写单寄存器出错，原始码 6，异常码 16#06 从站忙
 *   从站忙属告警级，可原样重试，短退避后再发即可，不必重启总线
 *   异常码 16#07 落在规范定义的编号空隙里，按未定义处理，故障级且有效性为假
 *============================================================================*)

FUNCTION FC_DL_ModbusExceptionParse : BOOL
VAR_INPUT
    uFuncCode : USINT;        // 响应功能码原值，最高位置位表示异常帧 [位串] / Raw response function code, top bit set means exception
    uExcCode  : USINT;        // 异常码，仅在异常帧有效 [代码] / Exception code, valid only on exception frames
END_VAR
VAR_OUTPUT
    bIsException : BOOL;                  // 是异常帧为真 / Exception frame detected
    nOrigFunc    : INT;                   // 原始功能码，去掉最高位后的值，0 表示非法 [代码] / Original function code without the top bit
    sExcName     : STRING(40);            // 异常码中文名，未定义码给「未定义异常码」 [文本] / Chinese name of the exception code
    eSeverity    : E_DL_ModbusExcSeverity; // 严重度分级，驱动上层重试策略 / Severity class driving the retry policy
    bRetryable   : BOOL;                  // 可原样重试为真 / Safe to retry unchanged
    uErrorId     : UDINT;                 // 事件码，0 表示无事件 / Event code, zero means none
    bValid       : BOOL;                  // 帧结构可解释为真 / Frame interpretable
END_VAR
VAR
    uFunc : USINT;            // 功能码快照，便于统一取位 [位串] / Function code snapshot
    uExc  : USINT;            // 异常码快照，便于分支判读 [代码] / Exception code snapshot
    nOrig : INT;              // 原始功能码中间量，先算后判 [代码] / Original code temporary
END_VAR
VAR CONSTANT
    DL_MB_EXC_BIT  : USINT := 16#80;   // 异常帧标志位，功能码最高位 [位串] / Exception flag bit, the top bit of the function code
    DL_MB_FUNC_MASK : USINT := 16#7F;  // 功能码掩码，去掉异常帧标志 [位串] / Function code mask removing the flag bit
    DL_MB_EXC_MAX  : USINT := 16#0B;   // 规范定义的异常码上限，超出即视为不可解释帧 [代码] / Highest code defined by the specification
END_VAR

(*------------------------------------------------------------------------------
 * 段 1｜输出预置：任何路径下输出确定
 *      Pre-set outputs so that every path is deterministic
 *-----------------------------------------------------------------------------*)
FC_DL_ModbusExceptionParse := FALSE;
bIsException               := FALSE;
nOrigFunc                  := 0;
sExcName                   := '';
eSeverity                  := E_DL_ModbusExcSeverity.eInfo;
bRetryable                 := FALSE;
uErrorId                   := 16#0000_0000;
bValid                     := FALSE;

(*------------------------------------------------------------------------------
 * 段 2｜取快照与异常帧判定（边界 B1）：最高位为异常标志
 *      Snapshot the inputs and detect the exception flag in the top bit
 *-----------------------------------------------------------------------------*)
uFunc        := uFuncCode;
uExc         := uExcCode;
bIsException := (uFunc AND DL_MB_EXC_BIT) <> 0;

(*------------------------------------------------------------------------------
 * 段 3｜原始功能码解出（边界 B2）：掩掉标志位，为零视为帧不可解释
 *      Strip the flag bit, a zero result means the frame cannot be interpreted
 *-----------------------------------------------------------------------------*)
nOrig     := USINT_TO_INT(uFunc AND DL_MB_FUNC_MASK);
nOrigFunc := nOrig;
IF nOrig = 0 THEN
    uErrorId := 16#0001_0138;   // 功能码非法，无原始语义可判
    RETURN;
END_IF

(*------------------------------------------------------------------------------
 * 段 4｜正常响应出口（边界 B3）：非异常帧给正常文字与信息码后返回
 *      Normal response exit: report the healthy frame and return
 *-----------------------------------------------------------------------------*)
IF NOT bIsException THEN
    sExcName                  := '正常响应';
    eSeverity                 := E_DL_ModbusExcSeverity.eInfo;
    bRetryable                := FALSE;
    bValid                    := TRUE;
    uErrorId                  := 16#0001_0139;   // 本帧不是异常帧，属提示
    FC_DL_ModbusExceptionParse := TRUE;
    RETURN;
END_IF

(*------------------------------------------------------------------------------
 * 段 5｜异常码映射（边界 B4）：逐码定性，未定义码走兜底分支
 *      Exception code mapping, undefined codes fall through to the fallback branch
 *      分级口径：组态类与校验类为故障级不可重试；忙与网关类为告警级可重试
 *-----------------------------------------------------------------------------*)
CASE uExc OF

    16#01:
        sExcName    := '非法功能';
        eSeverity   := E_DL_ModbusExcSeverity.eFault;
        bRetryable  := FALSE;

    16#02:
        sExcName    := '非法数据地址';
        eSeverity   := E_DL_ModbusExcSeverity.eFault;
        bRetryable  := FALSE;

    16#03:
        sExcName    := '非法数据值';
        eSeverity   := E_DL_ModbusExcSeverity.eFault;
        bRetryable  := FALSE;

    16#04:
        sExcName    := '从站设备故障';
        eSeverity   := E_DL_ModbusExcSeverity.eFault;
        bRetryable  := TRUE;

    16#05:
        sExcName    := '确认处理中';
        eSeverity   := E_DL_ModbusExcSeverity.eWarn;
        bRetryable  := TRUE;

    16#06:
        sExcName    := '从站设备忙';
        eSeverity   := E_DL_ModbusExcSeverity.eWarn;
        bRetryable  := TRUE;

    16#08:
        sExcName    := '存储奇偶校验错';
        eSeverity   := E_DL_ModbusExcSeverity.eFault;
        bRetryable  := FALSE;

    16#0A:
        sExcName    := '网关路径不可用';
        eSeverity   := E_DL_ModbusExcSeverity.eWarn;
        bRetryable  := TRUE;

    16#0B:
        sExcName    := '网关目标设备无响应';
        eSeverity   := E_DL_ModbusExcSeverity.eWarn;
        bRetryable  := TRUE;

    ELSE
        (* 未定义码兜底：文字照给便于 HMI 显示，但有效性置假，不算解析成功 *)
        (* Undefined code fallback: still name it for the HMI, but never mark it valid *)
        IF uExc > DL_MB_EXC_MAX THEN
            sExcName := '未定义异常码（超出规范上限）';
        ELSE
            sExcName := '未定义异常码';
        END_IF
        eSeverity  := E_DL_ModbusExcSeverity.eFault;
        bRetryable := FALSE;
        uErrorId   := 16#0001_0138;   // 未定义异常码，不可解释

END_CASE

(*------------------------------------------------------------------------------
 * 段 6｜收口：无事件即解析成功，事件码为未定义码时保持无效
 *      Close out: only event free calls count as a successful interpretation
 *-----------------------------------------------------------------------------*)
IF uErrorId = 16#0000_0000 THEN
    bValid                     := TRUE;
    FC_DL_ModbusExceptionParse := TRUE;
END_IF
END_FUNCTION

(* ---- FC_DL_ModbusRtuFrameCheck.st ---- *)
(*
    FC_DL_ModbusRtuFrameCheck —— Modbus RTU 帧一致性校验
    ------------------------------------------------------------------
    分类      : DL_MathData / Protocol
    前缀      : FC_DL_
    版本      : 1.0.0
    溯源      : Modbus 应用协议规范的公开条款（RTU 帧结构、功能码、异常应答长度、
                广播语义）；本库 T1-3 只借「协议帧解析与校验独立成族」的分类事实；
                判定表组织、错误分级、枚举范围与码位 100% 自有；CRC 校验另有
                FC_DL_Crc16Modbus，本件不重算 CRC；clean-room 重写，未复制任何
                闭源厂商源码，参考实现仅限 MIT/Apache 许可
    平台      : 纯 IEC 61131-3，CODESYS V3.5+ / TwinCAT 3 / InoProShop 通用
    作者      : 道莅代码库 · PLC编程专家（R19）
    ------------------------------------------------------------------
    功能说明  : 对已收到的 RTU 帧做结构一致性校验，把「解析异常帧」补成「先验帧再解帧」。
                四路互校：① 总长与功能码声明长度是否匹配；② 字节数域与调用方声明的
                数量 uQty 是否自洽；③ 异常帧（功能码 bit7 = 1）长度必须恰为 5；
                ④ 广播地址 0 配读类功能码属站号组态错（只提示不阻断）。
                核心防御：① 长度闸先于任何数组索引，绝不越界读 auFrame；
                ② 异常帧直接走定长分支，不做字节数互校（异常帧无字节数域）；
                ③ 未纳入长度表的功能码只做长度域检查并置信息码，不猜、不阻断上层；
                ④ CASE 含 ELSE 兜底，平台越界写入的非法枚举值同样按未识别功能码处理。
                职责边界：CRC 归 FC_DL_Crc16Modbus，异常码语义归 FC_DL_ModbusExceptionParse。
    错误码    : 16#0001_040A 功能码未纳入长度校验表（eFcUnknown / 非法枚举），只做长度域检查——信息级，正常防御
                16#0001_040B 广播地址配读类功能码（疑似站号组态错，已放行）——信息级，正常防御
                16#0001_032D 帧长非法（< 4 或 > 256 字节），不索引缓冲区——故障级，返回 FALSE
                16#0001_032E 字节数域 / 帧长与声明的数量 uQty 不自洽——故障级，返回 FALSE
                16#0001_032F 异常帧（bit7 置位）长度不等于 5——故障级，返回 FALSE
    码位总账  : 16#0001_040A 用 / 16#0001_040B 用 ｜ 16#0001_032D 用 / 16#0001_032E 用 / 16#0001_032F 用
    状态机    : R6 标注 N/A —— 本组件为纯函数无顺序状态机，无 CASE 可写，非法状态不可能出现
                （本件内部的 CASE 是功能码分派，不是顺序状态机，且含 ELSE 兜底）
    采样约定  : 本件无定时器、无沿检测；一帧一到即校验，结论与任务周期无关。
    修订记录  : 2026-11-16 v1.0.0 首次入库（R19）
*)

(*
    枚举 : E_DL_ModbusFc —— Modbus 功能码（本文件为全库唯一属主）
    说明 : 只覆盖本件能判定长度的 8 个功能码（01/02/03/04/05/06/0F/10）；
           08 诊断、0B 等一律 eFcUnknown 交上层处理，本件不猜。
*)
TYPE E_DL_ModbusFc :
(
    eFcUnknown := 0,                          // 未纳入长度校验表的功能码 / function code outside the length table
    eFc01      := 1,                          // 读线圈（位读取）/ read coils, bit read
    eFc02      := 2,                          // 读离散输入（位读取）/ read discrete inputs, bit read
    eFc03      := 3,                          // 读保持寄存器（字读取）/ read holding registers, word read
    eFc04      := 4,                          // 读输入寄存器（字读取）/ read input registers, word read
    eFc05      := 5,                          // 写单个线圈（定长 8 字节）/ write single coil, fixed 8 bytes
    eFc06      := 6,                          // 写单个寄存器（定长 8 字节）/ write single register, fixed 8 bytes
    eFc0F      := 15,                         // 写多个线圈（请求含字节数域）/ write multiple coils, request carries a byte count field
    eFc10      := 16                          // 写多个寄存器（请求含字节数域）/ write multiple registers, request carries a byte count field
);
END_TYPE

FUNCTION FC_DL_ModbusRtuFrameCheck : BOOL
VAR_INPUT
    auFrame         : ARRAY[0..255] OF BYTE;  // 帧缓冲区，定长 256 字节 / frame buffer, fixed 256 bytes
    uLen            : UINT := 0;              // 实际收到长度 [字节]，范围 0~256 / received length [byte], range 0~256
    eFc             : E_DL_ModbusFc := eFcUnknown; // 调用方读到的功能码（低 7 位语义）/ function code read by the caller, low seven bits
    uQty            : UINT := 0;              // 调用方声明的寄存器数或线圈数 [个]，范围 0~125 / declared register or coil quantity [count], range 0~125
END_VAR
VAR_OUTPUT
    eErr            : UDINT;                  // 错误码，0=正常 / error id, 0=ok
    bError          : BOOL;                   // 故障标志，eErr 为故障级时 TRUE / error flag, TRUE on fault-level eErr
    bValid          : BOOL;                   // 校验结论是否可信（故障态 FALSE）/ conclusion trustworthy flag, FALSE on fault
    uByteCount      : UINT;                   // 帧内解析出的字节数域 [字节]，无该域的功能码回 0 / byte count field parsed from the frame [byte], zero when absent
    bIsException    : BOOL;                   // 该帧是异常应答帧 / the frame is an exception response
    bBroadcast      : BOOL;                   // 地址域为 0（广播）/ address field is zero, broadcast
END_VAR
VAR CONSTANT
    DL_RTU_MIN_LEN   : UINT := 4;             // 最短帧长度（地址 + 功能码 + CRC×2）[字节] / shortest frame, address plus function code plus two CRC bytes [byte]
    DL_RTU_MAX_LEN   : UINT := 256;           // 协议与缓冲区上限 [字节] / protocol and buffer upper bound [byte]
    DL_RTU_EXC_LEN   : UINT := 5;             // 异常应答帧定长 [字节] / fixed exception response length [byte]
    DL_RTU_FIX_LEN   : UINT := 8;             // 05/06 定长帧 [字节] / fixed frame length for 05 and 06 [byte]
    DL_RTU_QTY_FIX   : UINT := 1;             // 05/06 允许的数量值（恒为 1）[个] / allowed quantity for 05 and 06, always one [count]
    DL_RTU_WR_BASE   : UINT := 9;             // 0F/10 请求帧最小长度（含 1 字节字节数域）[字节] / minimum request length for 0F and 10 [byte]
    DL_RTU_LEN_BASE  : UINT := 5;             // 读类应答帧固定开销（地址 + 功能码 + 字节数 + CRC×2）[字节] / fixed read response overhead [byte]
    DL_RTU_FC_EXC_BIT : BYTE := 16#80;        // 异常帧标志位（功能码 bit7）/ exception flag bit in the function code [bit]
    DL_RTU_BYTE_ZERO : BYTE := 16#00;         // 字节零常量，避免裸字面量 / byte zero constant, avoids a bare literal
    DL_RTU_ADDR_BROADCAST : BYTE := 16#00;    // 广播地址值 / broadcast address value
    DL_RTU_IDX_ADDR  : UINT := 0;             // 地址域下标 [索引] / address field index [index]
    DL_RTU_IDX_FC    : UINT := 1;             // 功能码域下标 [索引] / function code field index [index]
    DL_RTU_IDX_CNT   : UINT := 2;             // 读类应答的字节数域下标 [索引] / byte count index of a read response [index]
    DL_RTU_IDX_WRCNT : UINT := 6;             // 写多请求的字节数域下标 [索引] / byte count index of a multiple write request [index]
    DL_RTU_BITS_PER_BYTE : UINT := 8;         // 每字节位数，位数量换算用 [bit/字节] / bits per byte, used by the bit quantity conversion [bit/byte]
    DL_RTU_WORD_BYTES : UINT := 2;            // 每寄存器字节数 [字节/个] / bytes per register [byte/count]
    DL_RTU_BIT_ROUND : UINT := 7;             // 位数量上取整加数 [无量纲] / rounding addend for the bit quantity [dimensionless]
    DL_RTU_ZERO      : UINT := 0;             // 零值常量，避免裸字面量 [无量纲] / zero constant, avoids a bare literal [dimensionless]
    DL_RTU_ONE       : UINT := 1;             // 一值常量，下界判定用 [无量纲] / one constant used by the lower bound test [dimensionless]
END_VAR
VAR
    uExpectLen      : UINT;                   // 期望帧长中间量 [字节] / expected frame length intermediate [byte]
    uExpectCnt      : UINT;                   // 期望字节数域中间量 [字节] / expected byte count intermediate [byte]
    bWriteFc        : BOOL;                   // 是否为写类功能码（05/06/0F/10）/ write class function code flag
    bReadFc         : BOOL;                   // 是否为读类功能码（01/02/03/04）/ read class function code flag
    bFrameOk        : BOOL;                   // 帧结构自洽结论中间量 / frame self-consistency conclusion intermediate
END_VAR

// 段 1｜返回值与错误状态预置 / segment 1, preset return value and error status
FC_DL_ModbusRtuFrameCheck := FALSE;           // 缺省判定不自洽 / default conclusion is not self-consistent
eErr := 0;                                    // 预置无错误 / preset no error
bError := FALSE;                              // 预置无故障 / preset no fault
bValid := FALSE;                              // 预置结论不可信，通过闸门后置位 / preset untrustworthy, set TRUE after the gates
uByteCount := DL_RTU_ZERO;                    // 字节数域先清零 / clear the byte count field
bIsException := FALSE;                        // 预置非异常帧 / preset not an exception frame
bBroadcast := FALSE;                          // 预置非广播 / preset not a broadcast
bFrameOk := FALSE;                            // 结论中间量清零 / clear the conclusion intermediate
bWriteFc := FALSE;                            // 写类标志清零 / clear the write class flag
bReadFc := FALSE;                             // 读类标志清零 / clear the read class flag

// 段 2｜长度闸（先判长度再索引数组，绝不越界）/ segment 2, length gate before any indexing
IF (uLen < DL_RTU_MIN_LEN) OR (uLen > DL_RTU_MAX_LEN) THEN
    eErr := 16#0001_032D;                     // 帧长非法故障码 / illegal frame length fault id
    bError := TRUE;                           // 置故障标志 / raise the error flag
    bValid := FALSE;                          // 结论不可信 / conclusion untrustworthy
    RETURN;                                   // 故障级提前返回，不索引缓冲区 / early return, the buffer is never indexed
END_IF

// 段 3｜地址域判定（长度已保证下标 0 合法）/ segment 3, address field evaluation
bBroadcast := auFrame[DL_RTU_IDX_ADDR] = DL_RTU_ADDR_BROADCAST; // 地址 0 即广播 / address zero means broadcast

// 段 4｜异常帧分支：长度必须恰为 5，且不再做字节数互校 / segment 4, exception branch
IF (auFrame[DL_RTU_IDX_FC] AND DL_RTU_FC_EXC_BIT) <> DL_RTU_BYTE_ZERO THEN
    bIsException := TRUE;                     // 标记异常应答帧 / flag the exception response
    IF uLen = DL_RTU_EXC_LEN THEN
        bValid := TRUE;                       // 异常帧定长合法，结论可信 / fixed length is legal, the conclusion is trustworthy
        FC_DL_ModbusRtuFrameCheck := TRUE;    // 帧结构自洽 / the frame is self-consistent
    ELSE
        eErr := 16#0001_032F;                 // 异常帧长度非法故障码 / illegal exception frame length fault id
        bError := TRUE;                       // 置故障标志 / raise the error flag
        bValid := FALSE;                      // 结论不可信 / conclusion untrustworthy
        FC_DL_ModbusRtuFrameCheck := FALSE;   // 明确判定不自洽 / conclude not self-consistent
    END_IF
    RETURN;                                   // 异常帧分支出口，无字节数域可校 / exception frames carry no byte count field
END_IF

// 段 5｜功能码分派（含 ELSE 兜底，非法枚举按未识别处理）/ segment 5, function code dispatch with ELSE fallback
CASE eFc OF
    eFc01, eFc02:
        bReadFc := TRUE;                      // 位读取类 / bit read class
        IF uQty < DL_RTU_ONE THEN
            eErr := 16#0001_032E;             // 数量为 0 与功能码语义矛盾 / a zero quantity contradicts the function code
            bError := TRUE;                   // 置故障标志 / raise the error flag
        ELSE
            uByteCount := auFrame[DL_RTU_IDX_CNT]; // 解析字节数域 / parse the byte count field
            uExpectCnt := (uQty + DL_RTU_BIT_ROUND) / DL_RTU_BITS_PER_BYTE; // 位数量上取整为字节数，整数式禁浮点 / round the bit quantity up to bytes with integer arithmetic
            uExpectLen := DL_RTU_LEN_BASE + uExpectCnt; // 应答帧期望长度 / expected response length
            IF (uByteCount = uExpectCnt) AND (uLen = uExpectLen) THEN
                bFrameOk := TRUE;             // 字节数域与帧长双向自洽 / both the byte count and the length agree
            ELSE
                eErr := 16#0001_032E;         // 字节数域或帧长不自洽 / byte count or length mismatch
                bError := TRUE;               // 置故障标志 / raise the error flag
            END_IF
        END_IF

    eFc03, eFc04:
        bReadFc := TRUE;                      // 字读取类 / word read class
        IF uQty < DL_RTU_ONE THEN
            eErr := 16#0001_032E;             // 数量为 0 与功能码语义矛盾 / a zero quantity contradicts the function code
            bError := TRUE;                   // 置故障标志 / raise the error flag
        ELSE
            uByteCount := auFrame[DL_RTU_IDX_CNT]; // 解析字节数域 / parse the byte count field
            uExpectCnt := uQty * DL_RTU_WORD_BYTES; // 每寄存器 2 字节 / two bytes per register
            uExpectLen := DL_RTU_LEN_BASE + uExpectCnt; // 应答帧期望长度 / expected response length
            IF (uByteCount = uExpectCnt) AND (uLen = uExpectLen) THEN
                bFrameOk := TRUE;             // 字节数域与帧长双向自洽 / both the byte count and the length agree
            ELSE
                eErr := 16#0001_032E;         // 字节数域或帧长不自洽 / byte count or length mismatch
                bError := TRUE;               // 置故障标志 / raise the error flag
            END_IF
        END_IF

    eFc05, eFc06:
        bWriteFc := TRUE;                     // 写单点类 / single write class
        IF (uQty = DL_RTU_QTY_FIX) AND (uLen = DL_RTU_FIX_LEN) THEN
            bFrameOk := TRUE;                 // 定长帧且数量为 1 / fixed length frame with a quantity of one
        ELSE
            eErr := 16#0001_032E;             // 定长或数量不合法 / fixed length or quantity violated
            bError := TRUE;                   // 置故障标志 / raise the error flag
        END_IF

    eFc0F:
        bWriteFc := TRUE;                     // 写多点线圈类 / multiple coil write class
        IF (uQty >= DL_RTU_ONE) AND (uLen >= DL_RTU_WR_BASE) THEN
            uByteCount := auFrame[DL_RTU_IDX_WRCNT]; // 长度闸在前，下标 6 安全 / the length gate ran first, index six is safe
            uExpectCnt := (uQty + DL_RTU_BIT_ROUND) / DL_RTU_BITS_PER_BYTE; // 线圈数量换算字节数 / coil quantity converted to bytes
            IF uByteCount = uExpectCnt THEN
                bFrameOk := TRUE;             // 字节数域与声明数量自洽 / byte count agrees with the declared quantity
            ELSE
                eErr := 16#0001_032E;         // 字节数域不自洽 / byte count mismatch
                bError := TRUE;               // 置故障标志 / raise the error flag
            END_IF
        ELSE
            eErr := 16#0001_032E;             // 帧长或数量不足以承载请求 / length or quantity cannot carry the request
            bError := TRUE;                   // 置故障标志 / raise the error flag
        END_IF

    eFc10:
        bWriteFc := TRUE;                     // 写多点寄存器类 / multiple register write class
        IF (uQty >= DL_RTU_ONE) AND (uLen >= DL_RTU_WR_BASE) THEN
            uByteCount := auFrame[DL_RTU_IDX_WRCNT]; // 长度闸在前，下标 6 安全 / the length gate ran first, index six is safe
            uExpectCnt := uQty * DL_RTU_WORD_BYTES; // 每寄存器 2 字节 / two bytes per register
            IF uByteCount = uExpectCnt THEN
                bFrameOk := TRUE;             // 字节数域与声明数量自洽 / byte count agrees with the declared quantity
            ELSE
                eErr := 16#0001_032E;         // 字节数域不自洽 / byte count mismatch
                bError := TRUE;               // 置故障标志 / raise the error flag
            END_IF
        ELSE
            eErr := 16#0001_032E;             // 帧长或数量不足以承载请求 / length or quantity cannot carry the request
            bError := TRUE;                   // 置故障标志 / raise the error flag
        END_IF

    eFcUnknown:
        bFrameOk := TRUE;                     // 未纳入长度表：只做长度域检查后放行 / outside the table, released after the length check
        eErr := 16#0001_040A;                 // 信息级：功能码未纳入校验表 / info level, function code outside the length table

ELSE
    bFrameOk := TRUE;                         // 非法枚举值同样放行，不阻断上层解析 / illegal enum values are released too, never block the caller
    eErr := 16#0001_040A;                     // 信息级：未识别功能码，与 eFcUnknown 同一语义 / info level, unidentified function code, same semantics as eFcUnknown
END_CASE

// 段 6｜广播读类提示（协议上无意义，几乎必是站号配错；只提示不阻断）/ segment 6, broadcast read hint
IF (NOT bError) AND bBroadcast AND bReadFc THEN
    eErr := 16#0001_040B;                     // 信息级：广播配读类，已放行 / info level, broadcast with a read class, released
END_IF

// 段 7｜发布结论（故障级优先，信息码永不置 bError）/ segment 7, publish the conclusion
IF bError THEN
    FC_DL_ModbusRtuFrameCheck := FALSE;       // 故障态判定不自洽 / a fault means the frame is not self-consistent
    bValid := FALSE;                          // 结论不可信 / conclusion untrustworthy
ELSE
    FC_DL_ModbusRtuFrameCheck := bFrameOk;    // 无故障时输出结构自洽结论 / publish the self-consistency conclusion when no fault is present
    bValid := TRUE;                           // 结论可信 / conclusion trustworthy
END_IF
END_FUNCTION

(* ---- FC_DL_NewtonRaphson.st ---- *)
(*
  ==================================================================
  组件名 Component  : FC_DL_NewtonRaphson
  分类   Category   : DL_MathData
  版本   Version    : 1.0.0
  功能   Purpose    : 一元非线性方程牛顿迭代求根。主入口以多项式系数
                      a0..a8（下标即 x 的幂次）为方程定义，Horner 法一次
                      遍历同时得 f(x) 与解析 f'(x)；若置 bUseNumDiff 则改走
                      迭代内前向差分求导，免解析导数。副入口 FC_DL_NewtonStep
                      承载函数指针不可用时的两入口范式：调用侧用两个自有 FC
                      分别算出 f 与 f'，再逐步喂入 NewtonStep 推进迭代。
  防死锁 Anti-deadlock:
                      一 迭代次数硬上限 DL_NR_ITER_CAP = 200，入参超限钳到上限，
                         小于 1 钳 1；
                      二 收敛容差双端钳定 1E-12 / 1E-1，防「永不达标空转」与
                         「未迭代即判收敛」；
                      三 导数绝对值小于 lrDerivEps 立即退出并置 eDerivZero；
                      四 迭代量或残差出非有限值立即退出并置 eNonFinite；
                      五 残差连续 DL_NR_STALL_CAP 次无改善判停滞退出（eNoRoot）；
                      六 单步位移限幅 ±DL_NR_STEP_MAX，防坏导数放大成越界跳变。
  溯源   Origin     : 牛顿-拉夫逊迭代为公开数值方法。来源标签 t2-1-lgf-math（函数库
                      数学件分类域）；本件 clean-room 实现，仅借鉴来源分类与参数域
                      组织，未复制任何闭源代码行。
  平台   Platform   : 纯 IEC 61131-3（LREAL / WHILE / ABS / 无私有库、无方言转换）
  作者   Author     : 道莅代码库 · PLC 编程专家（R55）
  ------------------------------------------------------------------
  输入契约 Input contract:
                      afCoef 为引用型入参，由调用方持有并绑定，容量固定 9 项；
                      高阶项系数填 0 即按低阶多项式自然退化，无需裁剪数组。
  输出契约 Output contract:
                      eStatus 六态互斥；bConverged 仅 eOk 拍为 TRUE；bError 在一切
                      非 eOk 状态为 TRUE（含 eMaxIter 未达成，供上层判据用）；
                      bValid 仅在「根值有限 且 收敛或停滞」时为 TRUE；
                      根值非有限时出口回退初值 lrX0，非有限值不穿透出口。
  修订记录 Revision  :
    2026-11-20  v1.0.0  R55 首版（批 1 · 序号 1）
  ==================================================================
*)

TYPE E_DL_NrStatus :
(
    eOk        := 0,    // 收敛：残差已达容差 / converged, residual within tolerance
    eMaxIter   := 10,   // 达迭代上限未收敛 / iteration cap reached without convergence
    eDerivZero := 20,   // 导数近零：牛顿方向不可用 / derivative near zero, direction unusable
    eNonFinite := 30,   // 迭代中出非有限值（发散）/ non-finite value during iteration, diverged
    eBadArg    := 40,   // 入参非法：系数全零或入参非有限 / illegal argument, zero polynomial or non-finite input
    eNoRoot    := 50    // 停滞：残差连续无改善 / stalled, residual stopped improving
);
END_TYPE

FUNCTION FC_DL_NewtonRaphson : LREAL
VAR_IN_OUT
    afCoef      : ARRAY[0..8] OF LREAL;      // 多项式系数 a0..a8，下标即 x 的幂次 [无量纲]，引用型入参由调用方绑定 / coefficients a0..a8, subscript is the power of x [dimensionless], reference parameter bound by caller
END_VAR
VAR_INPUT
    lrX0        : LREAL := 0.0;              // 迭代初值 [无量纲] / initial guess [dimensionless]
    lrTol       : LREAL := 1.0E-9;           // 残差收敛容差 [无量纲]，双端钳定 / residual tolerance [dimensionless], clamped both ends
    lrDerivEps  : LREAL := 1.0E-10;          // 导数近零阈值 [无量纲]，导子绝对值小于即退出 / derivative near-zero threshold [dimensionless]
    nMaxIterIn  : INT := 50;                 // 期望最大迭代次数 [次]，超硬上限被钳 / requested max iterations [count], hard capped
    bUseNumDiff : BOOL := FALSE;             // 真 = 迭代内前向差分求导，假 = 解析导数 / true for in-loop forward difference, false for analytic derivative
    lrDiffStep  : LREAL := 1.0E-6;           // 差分步长 [无量纲]，域 大于零 / forward difference step [dimensionless], domain greater than zero
END_VAR
VAR_OUTPUT
    eStatus     : E_DL_NrStatus := E_DL_NrStatus.eOk; // 求根结果状态 [枚举] / root finding status [enum]
    nIterUsed   : INT := 0;                  // 实际迭代次数 [次] / iterations actually used [count]
    lrResidual  : LREAL := 0.0;              // 末次残差绝对值 [无量纲] / last absolute residual [dimensionless]
    bConverged  : BOOL := FALSE;             // 是否收敛 [-] / converged flag
    bError      : BOOL := FALSE;             // 是否未达成（任何非 eOk 状态）[-] / not achieved flag for any non-ok status
    bValid      : BOOL := FALSE;             // 根值是否可交付使用 [-] / root deliverable flag
END_VAR
VAR
    lrX         : LREAL := 0.0;              // 当前迭代点 [无量纲] / current iterate [dimensionless]
    lrFx        : LREAL := 0.0;              // 当前函数值 f(x) [无量纲] / current function value [dimensionless]
    lrFxH       : LREAL := 0.0;              // 差分点上函数值 f(x+h) [无量纲] / function value at the difference point [dimensionless]
    lrDf        : LREAL := 0.0;              // 当前导数值 f'(x) [无量纲] / current derivative value [dimensionless]
    lrStep      : LREAL := 0.0;              // 本步位移量 [无量纲] / current Newton step [dimensionless]
    lrResPrev   : LREAL := 0.0;              // 上一轮残差绝对值，停滞判据用 [无量纲] / previous residual for stall detection [dimensionless]
    lrTolUse    : LREAL := 1.0E-9;           // 钳定后的实际容差 [无量纲] / clamped effective tolerance [dimensionless]
    lrEpsUse    : LREAL := 1.0E-10;          // 钳定后的实际导数阈值 [无量纲] / clamped effective derivative threshold [dimensionless]
    lrHUse      : LREAL := 1.0E-6;           // 钳定后的实际差分步长 [无量纲] / clamped effective difference step [dimensionless]
    nIdx        : INT := 0;                  // 系数下标游标，向下递减 [下标] / coefficient index cursor, decremented [index]
    nIter       : INT := 0;                  // 迭代计数 [次] / iteration counter [count]
    nMaxIter    : INT := 1;                  // 钳定后的迭代上限 [次] / clamped iteration cap [count]
    nStall      : INT := 0;                  // 残差无改善连续计数 [次] / consecutive no-improvement count [count]
    bLoop       : BOOL := FALSE;             // 迭代循环续行标志 [-] / loop continuation flag
    bFinite     : BOOL := FALSE;             // 根值有限性判定暂存 [-] / root finiteness latch
    bCoefNz     : BOOL := FALSE;             // 多项式非全零判定暂存 [-] / non-zero polynomial latch
END_VAR
VAR CONSTANT
    DL_NR_ORD       : INT := 8;              // 多项式最高幂次，等于系数数组上界 [幂次] / highest polynomial order, equals coefficient upper bound
    DL_NR_ITER_CAP  : INT := 200;            // 迭代次数硬上限，防死锁 [次] / hard iteration cap against deadlock [count]
    DL_NR_TOL_MIN   : LREAL := 1.0E-12;      // 容差下限，防永不达标空转 [无量纲] / tolerance lower bound [dimensionless]
    DL_NR_TOL_MAX   : LREAL := 1.0E-1;       // 容差上限，防未迭代即判收敛 [无量纲] / tolerance upper bound [dimensionless]
    DL_NR_EPS_MIN   : LREAL := 1.0E-15;      // 导数阈值下限，防零阈致除零 [无量纲] / derivative threshold lower bound [dimensionless]
    DL_NR_STALL_CAP : INT := 5;              // 残差无改善连续次数上限 [次] / stall count cap [count]
    DL_NR_STEP_MAX  : LREAL := 1.0E9;        // 单步位移绝对上限 [无量纲] / single step absolute cap [dimensionless]
    DL_NR_H_MIN     : LREAL := 1.0E-9;       // 差分步长下限 [无量纲] / difference step lower bound [dimensionless]
    DL_NR_H_MAX     : LREAL := 1.0E-1;       // 差分步长上限 [无量纲] / difference step upper bound [dimensionless]
END_VAR

// 段 1｜返回值与错误状态预置，任何早退路径不留脏码 / segment 1, preset return value and error states, no dirty code on any early exit
FC_DL_NewtonRaphson := lrX0; // 返回值预置初值，非有限根时即以此值出口 / preset return to the initial guess, also the fallback when the root is non-finite
eStatus    := E_DL_NrStatus.eOk; // 状态预置收敛，后续按判定改写 / preset status to converged, rewritten by the following gates
nIterUsed  := 0; // 迭代计数出口预置零 / preset iteration count outlet to zero
lrResidual := 0.0; // 残差出口预置零 / preset residual outlet to zero
bConverged := FALSE; // 收敛标志预置假 / preset converged flag to false
bError     := FALSE; // 错误标志预置假 / preset error flag to false
bValid     := FALSE; // 有效标志预置假 / preset valid flag to false
lrX        := lrX0; // 迭代点从初值起步 / start the iterate from the initial guess

// 段 2｜入参域闸：容差双端钳定、迭代上限钳定、差分步长钳定、初值有限性 / segment 2, argument domain gate for tolerance, iteration cap, difference step and initial guess finiteness
lrTolUse := lrTol; // 容差默认直通 / tolerance passes through by default
IF lrTolUse <> lrTolUse THEN // 自反判 NaN / self-inequality detects NaN
    lrTolUse := DL_NR_TOL_MIN; // NaN 回落下限 / NaN falls back to the lower bound
END_IF
IF lrTolUse < DL_NR_TOL_MIN THEN // 容差过小 / tolerance too small
    lrTolUse := DL_NR_TOL_MIN; // 抬到下限，防永不达标空转 / raised to the lower bound against endless spinning
ELSIF lrTolUse > DL_NR_TOL_MAX THEN // 容差过大 / tolerance too large
    lrTolUse := DL_NR_TOL_MAX; // 压到上限，防未迭代即判收敛 / pressed to the upper bound against premature convergence
END_IF

lrEpsUse := lrDerivEps; // 导数阈值默认直通 / derivative threshold passes through by default
IF lrEpsUse <> lrEpsUse THEN // 自反判 NaN / self-inequality detects NaN
    lrEpsUse := DL_NR_EPS_MIN; // NaN 回落下限 / NaN falls back to the lower bound
END_IF
IF lrEpsUse < DL_NR_EPS_MIN THEN // 阈值过小 / threshold too small
    lrEpsUse := DL_NR_EPS_MIN; // 抬到下限，防除子近零 / raised against a near-zero divisor
ELSIF lrEpsUse > 1.0E-3 THEN // 阈值过大 / threshold too large
    lrEpsUse := 1.0E-3; // 压到 1E-3，防正常导数被误判近零 / pressed to 1E-3 against false near-zero verdicts
END_IF

lrHUse := lrDiffStep; // 差分步长默认直通 / difference step passes through by default
IF lrHUse <> lrHUse THEN // 自反判 NaN / self-inequality detects NaN
    lrHUse := 1.0E-6; // NaN 回落默认步长 / NaN falls back to the default step
END_IF
IF lrHUse < DL_NR_H_MIN THEN // 步长过小 / step too small
    lrHUse := DL_NR_H_MIN; // 抬到下限，防差分除子近零 / raised against a near-zero difference divisor
ELSIF lrHUse > DL_NR_H_MAX THEN // 步长过大 / step too large
    lrHUse := DL_NR_H_MAX; // 压到上限，防差分失真 / pressed against difference distortion
END_IF

nMaxIter := nMaxIterIn; // 迭代上限默认直通 / iteration cap passes through by default
IF nMaxIter < 1 THEN // 上限非法 / illegal cap
    nMaxIter := 1; // 钳到最少一次 / clamped to at least one iteration
ELSIF nMaxIter > DL_NR_ITER_CAP THEN // 上限越硬顶 / cap above the hard ceiling
    nMaxIter := DL_NR_ITER_CAP; // 钳到硬上限，防死锁 / clamped to the hard ceiling against deadlock
END_IF

// 段 3｜初值与系数有限性闸：非有限即判入参非法，不进迭代 / segment 3, finiteness gate on the initial guess and coefficients, illegal arguments never enter the loop
IF (lrX0 <> lrX0) OR ((lrX0 - lrX0) <> (lrX0 - lrX0)) THEN // 初值 NaN 或无穷 / initial guess is NaN or infinity
    eStatus := E_DL_NrStatus.eBadArg; // 入参非法 / illegal argument
    bError  := TRUE; // 置错误标志 / raise error flag
    bValid  := FALSE; // 出口不可用 / outlet unusable
    nIterUsed := 0; // 零次迭代 / zero iterations executed
    RETURN; // 早退，返回预置初值 / early exit with the preset initial guess
END_IF

bCoefNz := FALSE; // 多项式非全零标志预置假 / preset non-zero polynomial flag to false
nIdx := 0; // 下标游标归零 / reset the index cursor
WHILE nIdx <= DL_NR_ORD DO // 系数有限性与非全零双重扫查 / dual sweep for coefficient finiteness and non-zero content
    IF (afCoef[nIdx] <> afCoef[nIdx]) OR ((afCoef[nIdx] - afCoef[nIdx]) <> (afCoef[nIdx] - afCoef[nIdx])) THEN // 单项非有限 / single coefficient non-finite
        eStatus := E_DL_NrStatus.eBadArg; // 入参非法 / illegal argument
        bError  := TRUE; // 置错误标志 / raise error flag
        bValid  := FALSE; // 出口不可用 / outlet unusable
        RETURN; // 早退，返回预置初值 / early exit with the preset initial guess
    END_IF
    IF ABS(afCoef[nIdx]) > 0.0 THEN // 存在非零系数 / a non-zero coefficient exists
        bCoefNz := TRUE; // 置非全零标志 / raise the non-zero flag
    END_IF
    nIdx := nIdx + 1; // 游标递增，上界由 8 约束 / increment the cursor, upper bound fixed by eight
END_WHILE
IF NOT bCoefNz THEN // 全零多项式，任何点都是根 / zero polynomial, every point is a root
    eStatus := E_DL_NrStatus.eBadArg; // 入参非法，无求根意义 / illegal argument, root finding is meaningless
    bError  := TRUE; // 置错误标志 / raise error flag
    bValid  := FALSE; // 出口不可用 / outlet unusable
    RETURN; // 早退，返回预置初值 / early exit with the preset initial guess
END_IF

// 段 4｜牛顿迭代主循环：每轮先求值求导，再四级出口闸（收敛 / 导数近零 / 非有限 / 停滞）/ segment 4, Newton main loop with four exit gates per round
nIter    := 0; // 迭代计数清零 / reset the iteration counter
nStall   := 0; // 停滞计数清零 / reset the stall counter
lrResPrev := 0.0; // 残差快照清零 / reset the residual snapshot
bLoop    := TRUE; // 循环续行标志置真 / arm the loop continuation flag
WHILE bLoop AND (nIter < nMaxIter) DO // 循环条件含硬上限，双保险 / loop condition carries the hard cap as a second safety
    nIter := nIter + 1; // 迭代计数递增 / increment the iteration counter

    // 段 4.1｜Horner 同步求 f(x) 与解析 f'(x)，单遍复杂度 O(n) / segment 4.1, Horner yields both value and analytic derivative in one pass
    lrFx := afCoef[DL_NR_ORD]; // 从最高幂次系数起步 / start from the highest order coefficient
    lrDf := 0.0; // 导数累加器清零 / reset the derivative accumulator
    nIdx := DL_NR_ORD - 1; // 从次高幂次开始递减 / start one order below the highest
    WHILE nIdx >= 0 DO // 显式递减，规避负步进 FOR 的可移植风险 / explicit decrement avoids the portability risk of negative-step FOR
        lrDf := lrDf * lrX + lrFx; // 导数 Horner 递推 / derivative Horner recursion
        lrFx := lrFx * lrX + afCoef[nIdx]; // 函数值 Horner 递推 / value Horner recursion
        nIdx := nIdx - 1; // 游标递减 / decrement the cursor
    END_WHILE

    // 段 4.2｜差分模式覆盖解析导数（外部两入口不可用时的替代通路）/ segment 4.2, difference mode overrides the analytic derivative as the fallback path
    IF bUseNumDiff THEN // 差分模式生效 / difference mode active
        lrFxH := afCoef[DL_NR_ORD]; // 差分点求值从最高幂次系数起步 / difference point evaluation starts from the highest coefficient
        nIdx  := DL_NR_ORD - 1; // 差分求值下标重新起步 / restart the index cursor for the shifted evaluation
        WHILE nIdx >= 0 DO // 差分点同构 Horner / identical Horner at the shifted point
            lrFxH := lrFxH * (lrX + lrHUse) + afCoef[nIdx]; // 以 x + h 为自变量求值 / evaluate at x plus h
            nIdx  := nIdx - 1; // 游标递减 / decrement the cursor
        END_WHILE
        lrDf := (lrFxH - lrFx) / lrHUse; // 前向差分导数，除子已钳定大于零 / forward difference derivative, divisor proven positive
    END_IF

    // 段 4.3｜非有限闸：函数值或导数非有限即判发散退出，出口保持上拍值 / segment 4.3, non-finite gate, exit on divergence and keep the last healthy outlet
    IF (lrFx <> lrFx) OR ((lrFx - lrFx) <> (lrFx - lrFx)) OR (lrDf <> lrDf) OR ((lrDf - lrDf) <> (lrDf - lrDf)) THEN // 值或导数 NaN 或无穷 / value or derivative is NaN or infinity
        eStatus := E_DL_NrStatus.eNonFinite; // 发散退出 / diverged exit
        bLoop   := FALSE; // 终止循环 / terminate the loop
    ELSE
        lrResidual := ABS(lrFx); // 残差取绝对值 / residual as an absolute value
        IF lrResidual <= lrTolUse THEN // 收敛出口 / convergence exit
            bConverged := TRUE; // 置收敛标志 / raise the converged flag
            eStatus    := E_DL_NrStatus.eOk; // 状态记收敛 / record the converged status
            bLoop      := FALSE; // 终止循环 / terminate the loop
        ELSIF ABS(lrDf) < lrEpsUse THEN // 导数近零出口 / derivative near-zero exit
            eStatus := E_DL_NrStatus.eDerivZero; // 方向不可用 / direction unusable
            bLoop   := FALSE; // 终止循环 / terminate the loop
        ELSE
            lrStep := -lrFx / lrDf; // 牛顿位移，除子绝对值已证不小于阈值 / Newton step, divisor magnitude proven not below the threshold
            IF lrStep > DL_NR_STEP_MAX THEN // 正越界 / positive overflow
                lrStep := DL_NR_STEP_MAX; // 上钳到步长上限 / clamp to the positive step cap
            ELSIF lrStep < -DL_NR_STEP_MAX THEN // 负越界 / negative overflow
                lrStep := -DL_NR_STEP_MAX; // 下钳到步长上限 / clamp to the negative step cap
            END_IF
            lrX := lrX + lrStep; // 推进迭代点 / advance the iterate
            IF (lrX <> lrX) OR ((lrX - lrX) <> (lrX - lrX)) THEN // 新点非有限 / new point non-finite
                eStatus := E_DL_NrStatus.eNonFinite; // 发散退出 / diverged exit
                bLoop   := FALSE; // 终止循环 / terminate the loop
            ELSE
                IF (nIter > 1) AND (lrResidual >= lrResPrev * 0.999) THEN // 残差无实质改善 / residual did not improve materially
                    nStall := nStall + 1; // 停滞计数递增 / increment the stall counter
                ELSE
                    nStall := 0; // 有改善则清零 / clear on improvement
                END_IF
                lrResPrev := lrResidual; // 更新残差快照 / refresh the residual snapshot
                IF nStall >= DL_NR_STALL_CAP THEN // 停滞达上限 / stall count reached the cap
                    eStatus := E_DL_NrStatus.eNoRoot; // 判停滞退出 / stalled exit
                    bLoop   := FALSE; // 终止循环 / terminate the loop
                END_IF
            END_IF
        END_IF
    END_IF
END_WHILE

// 段 5｜循环自然结束仍未收敛者判达上限（eOk 以外的既有状态不覆盖）/ segment 5, a natural loop end without convergence is an iteration-cap verdict, existing non-ok statuses are preserved
IF bLoop AND (NOT bConverged) AND (eStatus = E_DL_NrStatus.eOk) THEN // 循环用完次数且无其它出口 / iterations exhausted with no other exit
    eStatus := E_DL_NrStatus.eMaxIter; // 达上限未收敛 / cap reached without convergence
END_IF

// 段 6｜统一出口：有限性闸 + 根值交付 + 标志落定 / segment 6, unified outlet with finiteness gate, root delivery and flag settling
nIterUsed := nIter; // 迭代次数出口落定 / settle the iteration count outlet
bFinite   := (lrX = lrX) AND ((lrX - lrX) = (lrX - lrX)); // 根值有限性判定，NaN 用自反、无穷用差值自减 / root finiteness by self-inequality for NaN and self-difference for infinity
IF bFinite THEN // 根值有限 / root is finite
    FC_DL_NewtonRaphson := lrX; // 交付根值 / deliver the root
    bValid := bConverged OR (eStatus = E_DL_NrStatus.eNoRoot); // 收敛或停滞的有限根可交付，其余状态仅供诊断 / finite roots from convergence or stall are deliverable, other statuses are diagnostic only
ELSE
    FC_DL_NewtonRaphson := lrX0; // 非有限：退回初值，非有限值不穿透出口 / non-finite, fall back to the initial guess so nothing non-finite passes the outlet
    bValid := FALSE; // 出口不可用 / outlet unusable
END_IF
bError := NOT (eStatus = E_DL_NrStatus.eOk); // 任何非收敛状态均置错误标志，供上层判据 / any non-converged status raises the error flag for the upper layer
END_FUNCTION

(*
  ------------------------------------------------------------------
  FC_DL_NewtonStep —— 两入口推进单步（函数指针不可用时的配套入口）
  ------------------------------------------------------------------
  功能说明  : 供调用侧「两入口」使用：调用侧分别用自有 FC 算出 f(x) 与 f'(x)，
              把两个数值与本拍迭代点喂入本 FC，得到推进后的下一个迭代点。
              本 FC 无内部状态，调用侧持有循环与迭代上限（自身需另设硬上限）。
              与主入口同一套出口闸：值/导数非有限、导数近零、位移越界均拒绝推进。
  输出契约  : lrNextX 在拒推拍保持 lrX（不推进，等价于出口保持上拍值）；
              bStepOk 仅在本次推进合法时为 TRUE；eStatus 复用同一枚举。
  修订记录  : 2026-11-20 v1.0.0 R55 首版（与主入口同文件交付）
*)
FUNCTION FC_DL_NewtonStep : LREAL
VAR_INPUT
    lrX         : LREAL := 0.0;              // 当前迭代点 [无量纲] / current iterate [dimensionless]
    lrF         : LREAL := 0.0;              // 外部入口一算出的函数值 f(x) [无量纲] / function value from external entry one [dimensionless]
    lrDf        : LREAL := 0.0;              // 外部入口二算出的导数值 f'(x) [无量纲] / derivative value from external entry two [dimensionless]
    lrDerivEps  : LREAL := 1.0E-10;          // 导数近零阈值 [无量纲] / derivative near-zero threshold [dimensionless]
    lrStepMax   : LREAL := 1.0E9;            // 单步位移绝对上限 [无量纲] / single step absolute cap [dimensionless]
END_VAR
VAR_OUTPUT
    bStepOk     : BOOL := FALSE;             // 本次推进是否合法 [-] / whether this advance is legal
    eStatus     : E_DL_NrStatus := E_DL_NrStatus.eOk; // 推进结果状态 [枚举] / advance status [enum]
END_VAR
VAR
    lrStep      : LREAL := 0.0;              // 本步位移量 [无量纲] / current step [dimensionless]
    lrEps       : LREAL := 1.0E-10;          // 钳定后的导数阈值 [无量纲] / clamped derivative threshold [dimensionless]
    lrCap       : LREAL := 1.0E9;            // 钳定后的位移上限 [无量纲] / clamped step cap [dimensionless]
END_VAR
VAR CONSTANT
    DL_NS_EPS_MIN : LREAL := 1.0E-15;        // 导数阈值下限，防零阈致除零 [无量纲] / derivative threshold lower bound against division by zero
    DL_NS_CAP_MIN : LREAL := 1.0E-3;         // 位移上限下限，防零上限锁死推进 [无量纲] / step cap lower bound against a locked advance
END_VAR

// 段 1｜出口预置：默认不推进，保持传入迭代点 / segment 1, preset the outlet to no advance, keeping the incoming iterate
FC_DL_NewtonStep := lrX; // 拒推拍返回原点 / return the incoming point when the advance is rejected
bStepOk := FALSE; // 推进标志预置假 / preset the advance flag to false
eStatus := E_DL_NrStatus.eOk; // 状态预置收敛 / preset status to converged

// 段 2｜阈值与上限域闸 / segment 2, domain gate for the threshold and the cap
lrEps := lrDerivEps; // 阈值默认直通 / threshold passes through by default
IF lrEps <> lrEps THEN // 自反判 NaN / self-inequality detects NaN
    lrEps := DL_NS_EPS_MIN; // NaN 回落下限 / NaN falls back to the lower bound
END_IF
IF lrEps < DL_NS_EPS_MIN THEN // 阈值过小 / threshold too small
    lrEps := DL_NS_EPS_MIN; // 抬到下限 / raised to the lower bound
END_IF
lrCap := lrStepMax; // 位移上限默认直通 / step cap passes through by default
IF lrCap <> lrCap THEN // 自反判 NaN / self-inequality detects NaN
    lrCap := 1.0E9; // NaN 回落默认上限 / NaN falls back to the default cap
END_IF
IF lrCap < DL_NS_CAP_MIN THEN // 上限过小 / cap too small
    lrCap := DL_NS_CAP_MIN; // 抬到下限，防推进被锁死 / raised against a locked advance
END_IF

// 段 3｜三入口有限性闸：任一项非有限即拒绝推进 / segment 3, finiteness gate on all three inputs, any non-finite term rejects the advance
IF (lrX <> lrX) OR ((lrX - lrX) <> (lrX - lrX)) OR (lrF <> lrF) OR ((lrF - lrF) <> (lrF - lrF)) OR (lrDf <> lrDf) OR ((lrDf - lrDf) <> (lrDf - lrDf)) THEN // 任一项 NaN 或无穷 / any term is NaN or infinity
    eStatus := E_DL_NrStatus.eNonFinite; // 非有限拒绝 / rejected as non-finite
    RETURN; // 早退，出口保持传入点 / early exit with the outlet held at the incoming point
END_IF

// 段 4｜导数闸与位移限幅 / segment 4, derivative gate and step clamp
IF ABS(lrDf) < lrEps THEN // 导数近零 / derivative near zero
    eStatus := E_DL_NrStatus.eDerivZero; // 方向不可用 / direction unusable
    RETURN; // 早退，出口保持传入点 / early exit with the outlet held at the incoming point
END_IF
lrStep := -lrF / lrDf; // 牛顿位移，除子绝对值已证不小于阈值 / Newton step, divisor magnitude proven not below the threshold
IF lrStep > lrCap THEN // 正越界 / positive overflow
    lrStep := lrCap; // 上钳 / clamp upward
ELSIF lrStep < -lrCap THEN // 负越界 / negative overflow
    lrStep := -lrCap; // 下钳 / clamp downward
END_IF

// 段 5｜推进与结果有限性复检 / segment 5, advance and finiteness recheck
FC_DL_NewtonStep := lrX + lrStep; // 推进到下一个迭代点 / advance to the next iterate
IF (FC_DL_NewtonStep <> FC_DL_NewtonStep) OR ((FC_DL_NewtonStep - FC_DL_NewtonStep) <> (FC_DL_NewtonStep - FC_DL_NewtonStep)) THEN // 新点非有限 / new point non-finite
    eStatus := E_DL_NrStatus.eNonFinite; // 判发散 / diverged verdict
    FC_DL_NewtonStep := lrX; // 退回原迭代点 / fall back to the incoming iterate
    bStepOk := FALSE; // 推进标志保持假 / advance flag stays false
    RETURN; // 早退 / early exit
END_IF
bStepOk := TRUE; // 推进合法 / the advance is legal
eStatus := E_DL_NrStatus.eOk; // 状态记正常 / record the normal status
END_FUNCTION
